FUNCTION FC 911 : VOID
TITLE =NEW FC911 (was FC1011) - Conveyors - Clearing Function
//New Order Sequence
//v0.1 2026-11-19: hold released at clearing start (FP M283.4); S3.2 lamp steady
//while held / blinking when ready; S3.2 held 3s releases the hold (T140).
//v0.2 2026-11-19: C10 empty proof added up over several runs (MD284), time from
//Surface_Length_10 (no more waiting for the bottomer). T137 no longer used.
//v0.3 2026-11-19: C10 empty proof by ENCODER TRAVEL (PIW 334 direct), not time:
//travel >= Surface_Length_10 + 20 % with exit clear, added up (MD284, MW288).
//v0.4 2026-11-19: encoder steps < 0 or > 300 pulses/scan ignored (Ch5 restarts
//from 0 when its gate reopens, every 500 mS while clearing) - no false proof.
NAME : CLEARING
VERSION : 0.4


VAR_TEMP
  EMPTY_11 : BOOL ;	//Empty Conveyor 11
  EMPTY_21 : BOOL ;	//Empty Conveyor 21
  EMPTY_12_22 : BOOL ;	//Empty Conveyor 12 & 22
  EMPTY_13_23 : BOOL ;	//Empty Conveyor 13 & 23
  C10_EMPTY_TEST : BOOL ;
  CLEARING_ABORT : BOOL ;
  PROOF_P : DINT ;	//C10 Empty Proof Travel [Pulses]
  D_ENC : DINT ;	//Encoder Pulses This Scan
  ENC_W : INT ;	//Encoder Word PIW 334
END_VAR
BEGIN
NETWORK
TITLE =HMI Clearing Call

      A     "M 140.3";
      A     "HMI_DB".CLEARING_SSW_MAIN;
      =     "M 5.2";
//;
      L     8;
      A     "M 10.0";
      =     "HMI_DB".CLEARING_SSW_STATUS;
      JC    CLEA;

      L     0;

CLEA: T     "HMI_DB".CLEARING_FUNCTION;

      A     "M 10.0";
      FN    "FN 155.7";
      R     "HMI_DB".CLEARING_SSW_MAIN;
      R     "M 54.2";
//;
      A     "M 5.2";
      FP    "FP 147.4";
      AN    "B 10.7"; // C11 - Empty
      AN    "B 11.0"; // C12 - Empty
      AN    "B 11.1"; // C13 - Empty
      AN    "B 11.2"; // C13 - Empty
      AN    "B 15.4"; // C21 - Empty
      AN    "B 15.5"; // C22 - Empty
      AN    "B 15.6"; // C23 - Empty
      AN    "B 15.7"; // C23 - Empty
      S     "M 54.2"; // Empty C11...C23
NETWORK
TITLE =New Order Seq - First New Order Packet to Pivot Conveyor 10
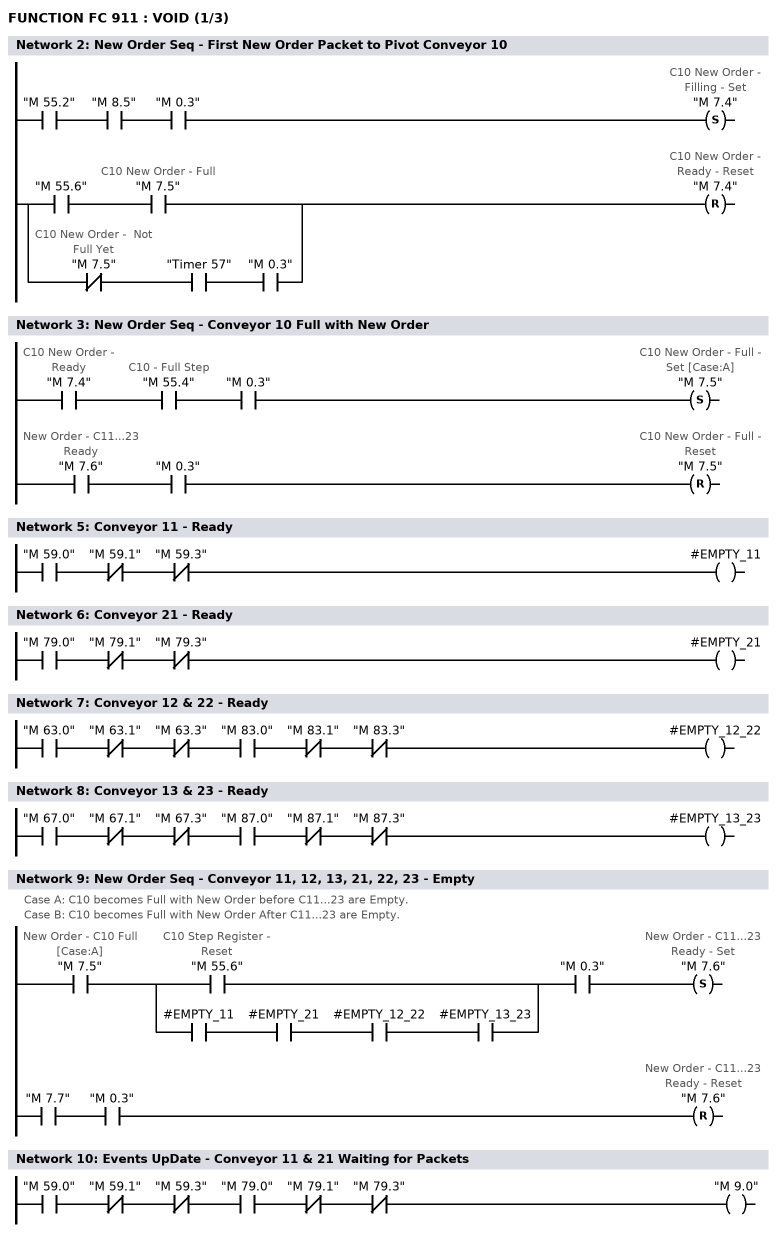

      A     "M 55.2";
      A     "M 8.5";
      A     "M 0.3";
      S     "M 7.4"; // C10 New Order - Filling - Set
//;
      A(    ;
      A     "M 55.6";
      A     "M 7.5"; // C10 New Order - Full
      O     ;
      AN    "M 7.5"; // C10 New Order -  Not Full Yet
      A     "Timer 57";
      A     "M 0.3";
      )     ;
      R     "M 7.4"; // C10 New Order - Ready - Reset
NETWORK
TITLE =New Order Seq - Conveyor 10 Full with New Order

      A     "M 7.4"; // C10 New Order - Ready
      A     "M 55.4"; // C10 - Full Step
      A     "M 0.3";
      S     "M 7.5"; // C10 New Order - Full - Set [Case:A]
//;
      A     "M 7.6"; // New Order - C11...23 Ready
      A     "M 0.3";
      R     "M 7.5"; // C10 New Order - Full - Reset
NETWORK
TITLE =New Order Seq
//New Order Seq - Waiting for the last Order Packets to Run out !


NETWORK
TITLE =Conveyor 11 - Ready

      A     "M 59.0";
      AN    "M 59.1";
      AN    "M 59.3";
      =     #EMPTY_11;
NETWORK
TITLE =Conveyor 21 - Ready

      A     "M 79.0";
      AN    "M 79.1";
      AN    "M 79.3";
      =     #EMPTY_21;
NETWORK
TITLE =Conveyor 12 & 22 - Ready

      A     "M 63.0";
      AN    "M 63.1";
      AN    "M 63.3";
      A     "M 83.0";
      AN    "M 83.1";
      AN    "M 83.3";
      =     #EMPTY_12_22;
NETWORK
TITLE =Conveyor 13 & 23 - Ready

      A     "M 67.0";
      AN    "M 67.1";
      AN    "M 67.3";
      A     "M 87.0";
      AN    "M 87.1";
      AN    "M 87.3";
      =     #EMPTY_13_23;
NETWORK
TITLE =New Order Seq - Conveyor 11, 12, 13, 21, 22, 23 - Empty
//Case A: C10 becomes Full with New Order before C11...23 are Empty.
//Case B: C10 becomes Full with New Order After C11...23 are Empty.
      A     "M 7.5"; // New Order - C10 Full [Case:A]
      A(    ;
      A     "M 55.6"; // C10 Step Register - Reset
      O     ;
      A     #EMPTY_11;
      A     #EMPTY_21;
      A     #EMPTY_12_22;
      A     #EMPTY_13_23;
      )     ;
      A     "M 0.3";
      S     "M 7.6"; // New Order - C11...23 Ready - Set
//;
      A     "M 7.7";
      A     "M 0.3";
      R     "M 7.6"; // New Order - C11...23 Ready - Reset
NETWORK
TITLE =Events UpDate - Conveyor 11 & 21 Waiting for Packets

      A     "M 59.0";
      AN    "M 59.1";
      AN    "M 59.3";
      A     "M 79.0";
      AN    "M 79.1";
      AN    "M 79.3";
      =     "M 9.0";
NETWORK
TITLE =New Order Seq - Conveyors 11, 21 - Empty
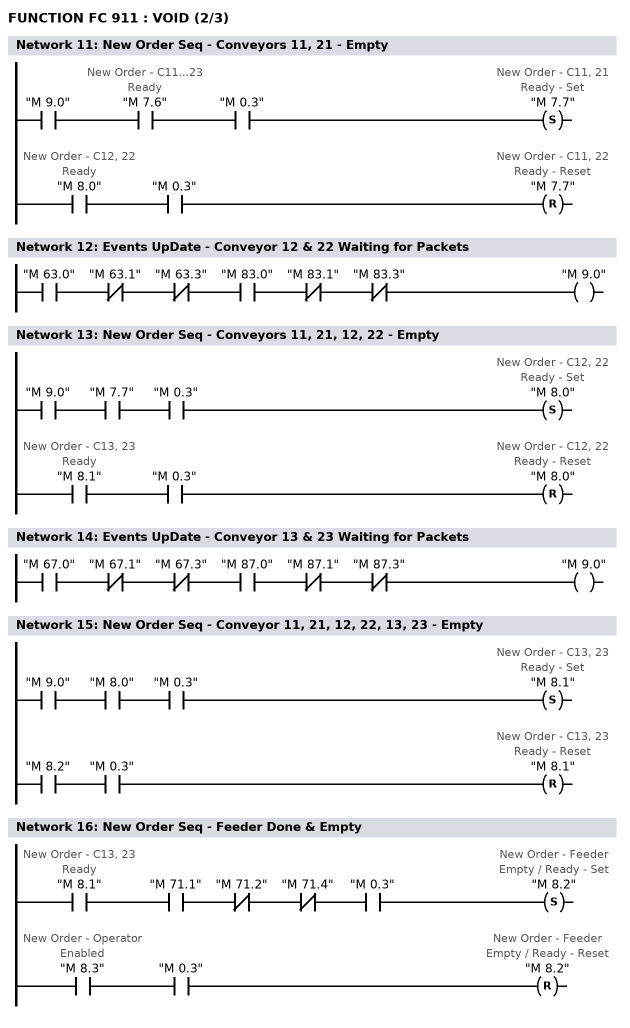

      A     "M 9.0";
      A     "M 7.6"; // New Order - C11...23 Ready
      A     "M 0.3";
      S     "M 7.7"; // New Order - C11, 21 Ready - Set
//;
      A     "M 8.0"; // New Order - C12, 22 Ready
      A     "M 0.3";
      R     "M 7.7"; // New Order - C11, 22 Ready - Reset
NETWORK
TITLE =Events UpDate - Conveyor 12 & 22 Waiting for Packets

      A     "M 63.0";
      AN    "M 63.1";
      AN    "M 63.3";
      A     "M 83.0";
      AN    "M 83.1";
      AN    "M 83.3";
      =     "M 9.0";
NETWORK
TITLE =New Order Seq - Conveyors 11, 21, 12, 22 - Empty

      A     "M 9.0";
      A     "M 7.7";
      A     "M 0.3";
      S     "M 8.0"; // New Order - C12, 22 Ready - Set
//;
      A     "M 8.1"; // New Order - C13, 23 Ready
      A     "M 0.3";
      R     "M 8.0"; // New Order - C12, 22 Ready - Reset
NETWORK
TITLE =Events UpDate - Conveyor 13 & 23 Waiting for Packets

      A     "M 67.0";
      AN    "M 67.1";
      AN    "M 67.3";
      A     "M 87.0";
      AN    "M 87.1";
      AN    "M 87.3";
      =     "M 9.0";
NETWORK
TITLE =New Order Seq - Conveyor 11, 21, 12, 22, 13, 23 - Empty

      A     "M 9.0";
      A     "M 8.0";
      A     "M 0.3";
      S     "M 8.1"; // New Order - C13, 23 Ready - Set
//;
      A     "M 8.2";
      A     "M 0.3";
      R     "M 8.1"; // New Order - C13, 23 Ready - Reset
NETWORK
TITLE =New Order Seq - Feeder Done & Empty

      A     "M 8.1"; // New Order - C13, 23 Ready
      A     "M 71.1";
      AN    "M 71.2";
      AN    "M 71.4";
      A     "M 0.3";
      S     "M 8.2"; // New Order - Feeder Empty / Ready - Set
//;
      A     "M 8.3"; // New Order - Operator Enabled
      A     "M 0.3";
      R     "M 8.2"; // New Order - Feeder Empty / Ready - Reset
NETWORK
TITLE =Conveyor 10 Clearing Enable after New Order
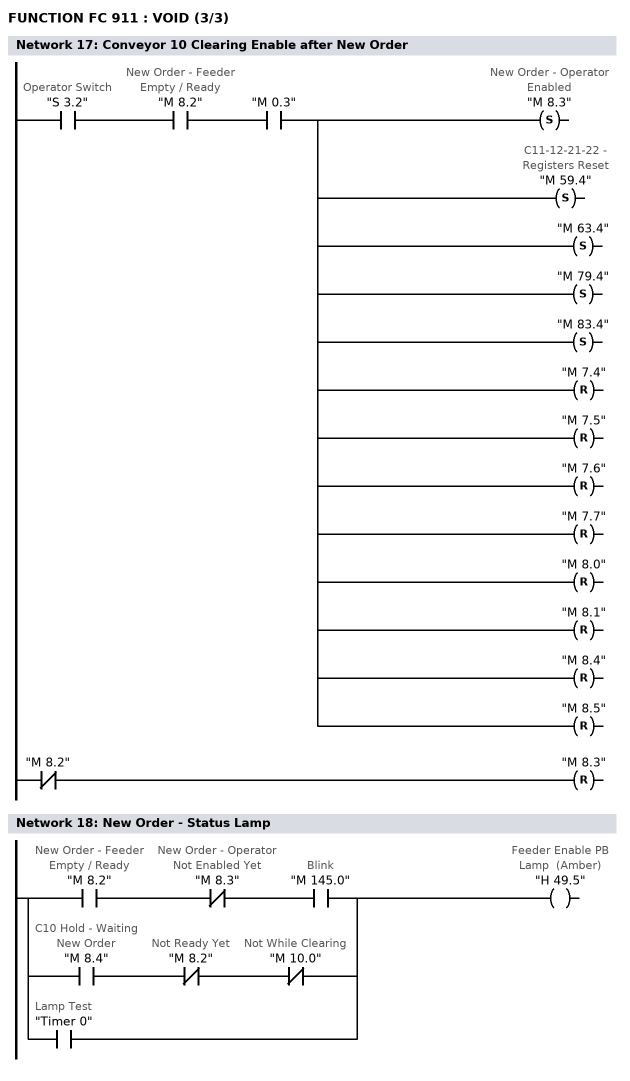

      A     "S 3.2"; // Operator Switch
      A     "M 8.2"; // New Order - Feeder Empty / Ready
      A     "M 0.3";
      S     "M 8.3"; // New Order - Operator Enabled
      S     "M 59.4"; // C11-12-21-22 - Registers Reset
      S     "M 63.4";
      S     "M 79.4";
      S     "M 83.4";
//;
      R     "M 7.4";
      R     "M 7.5";
      R     "M 7.6";
      R     "M 7.7";
      R     "M 8.0";
      R     "M 8.1";
      R     "M 8.4";
      R     "M 8.5";
//;
      ON    "M 8.2";
      R     "M 8.3";
NETWORK
TITLE =New Order - Status Lamp

//2026-11-19: BLINK = S3.2 can be pressed now (M8.2). STEADY = C10 held for the
//new order, not ready yet (M8.4 without M8.2) - before, the lamp stayed OFF.
      A(    ;
      A     "M 8.2"; // New Order - Feeder Empty / Ready
      AN    "M 8.3"; // New Order - Operator Not Enabled Yet
      A     "M 145.0"; // Blink
      )     ;
      O(    ;
      A     "M 8.4"; // C10 Hold - Waiting New Order
      AN    "M 8.2"; // Not Ready Yet
      AN    "M 10.0"; // Not While Clearing
      )     ;
      O     "Timer 0"; // Lamp Test
      =     "H 49.5"; // Feeder Enable PB Lamp  (Amber)
NETWORK
TITLE =S3.2 Held 3s - Release the Hold (Sequence Not Complete)
//2026-11-19: Before, S3.2 only worked with M8.2 (whole new-order chain done).
//If the chain got stuck, the TS waited with no way out but SIGNAL/F4.
//S3.2 held 3s releases the hold only (C11...C22 steps NOT reset: they may
//still carry the previous order).

      A     "S 3.2"; // Operator PB
      A     "M 8.4"; // C10 Hold Active
      AN    "M 10.0"; // Not While Clearing
      L     S5T#3S;
      SD    T    140; // Hold 3s (Free Timer)
//;
      A     T    140;
      A     "M 0.3";
      JCN   S321;

      R     "M 7.4";
      R     "M 7.5";
      R     "M 7.6";
      R     "M 7.7";
      R     "M 8.0";
      R     "M 8.1";
      R     "M 8.2";
      R     "M 8.3";
      R     "M 8.4"; // C10 Hold - Released
      R     "M 8.5"; // Clearing Done - Reset

S321: NOP   0;
NETWORK
TITLE =Conveyors Clearing Blink
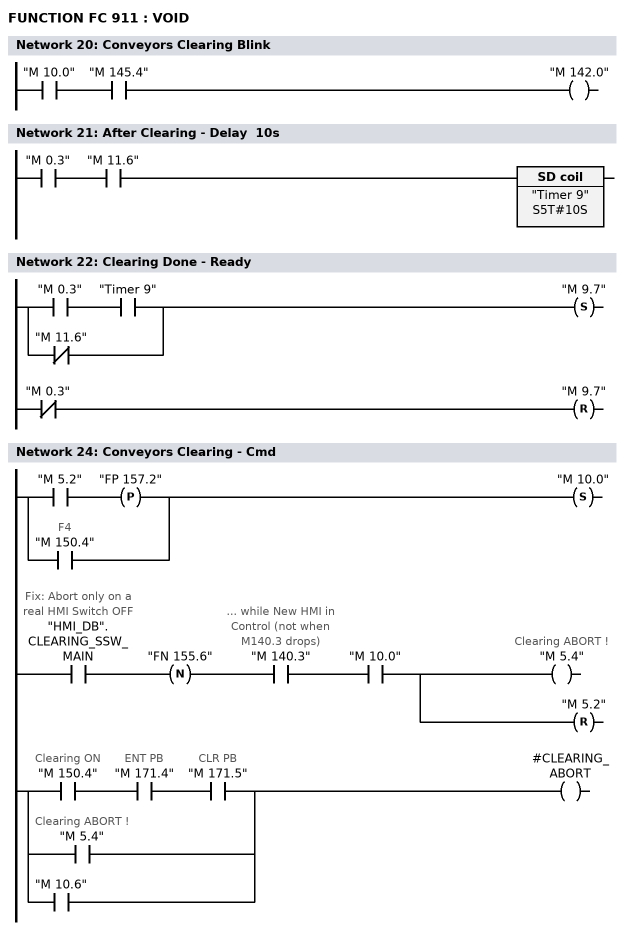

      A     "M 10.0";
      A     "M 145.4";
      =     "M 142.0";
NETWORK
TITLE =After Clearing - Delay  10s

      A     "M 0.3";
      A     "M 11.6";
      L     S5T#10S;
      SD    "Timer 9";
NETWORK
TITLE =Clearing Done - Ready

      A     "M 0.3";
      A     "Timer 9";
      ON    "M 11.6";
      S     "M 9.7";
//;
      ON    "M 0.3";
      R     "M 9.7";
NETWORK
TITLE =Clearing Command
//Clearing Command


NETWORK
TITLE =Conveyors Clearing - Cmd

      A(    ;
      A     "M 5.2";
      FP    "FP 157.2";
      O     ;
      A     "M 150.4"; // F4
      )     ;
      S     "M 10.0";
//;
      A     "HMI_DB".CLEARING_SSW_MAIN; // Fix: Abort only on a real HMI Switch OFF
      FN    "FN 155.6";
      A     "M 140.3"; // ... while New HMI in Control (not when M140.3 drops)
      A     "M 10.0";
      =     "M 5.4"; // Clearing ABORT !
      R     "M 5.2";
//;
      A(    ;
      A     "M 150.4"; // Clearing ON
      A     "M 171.4"; // ENT PB
      A     "M 171.5"; // CLR PB
      O     "M 5.4"; // Clearing ABORT !
      O     "M 10.6";
      )     ;
      =     #CLEARING_ABORT;
NETWORK
TITLE =Clearing Start - Release a Hold Left from the Previous Clearing
//Fix 2026-11-19: F4 pressed while C10 still held a new order (M8.4, S3.2 not
//pressed yet) -> C10 could not transfer, the clearing could never finish.
//F4 = clear everything: at every clearing start the hold and the new-order
//sequence are reset. They are set again when this clearing is done.

      A     "M 10.0"; // Clearing CMD
      FP    M    283.4; // Edge Memory (Free)
      JCN   CST1;

      R     "M 7.4";
      R     "M 7.5";
      R     "M 7.6";
      R     "M 7.7";
      R     "M 8.0";
      R     "M 8.1";
      R     "M 8.2";
      R     "M 8.3";
      R     "M 8.4"; // C10 Hold - Released
      R     "M 8.5"; // Clearing Done - Reset

CST1: NOP   0;
NETWORK
TITLE =Conveyors Clearing Conveyors 1,2,3,4 - TimeOut 30S
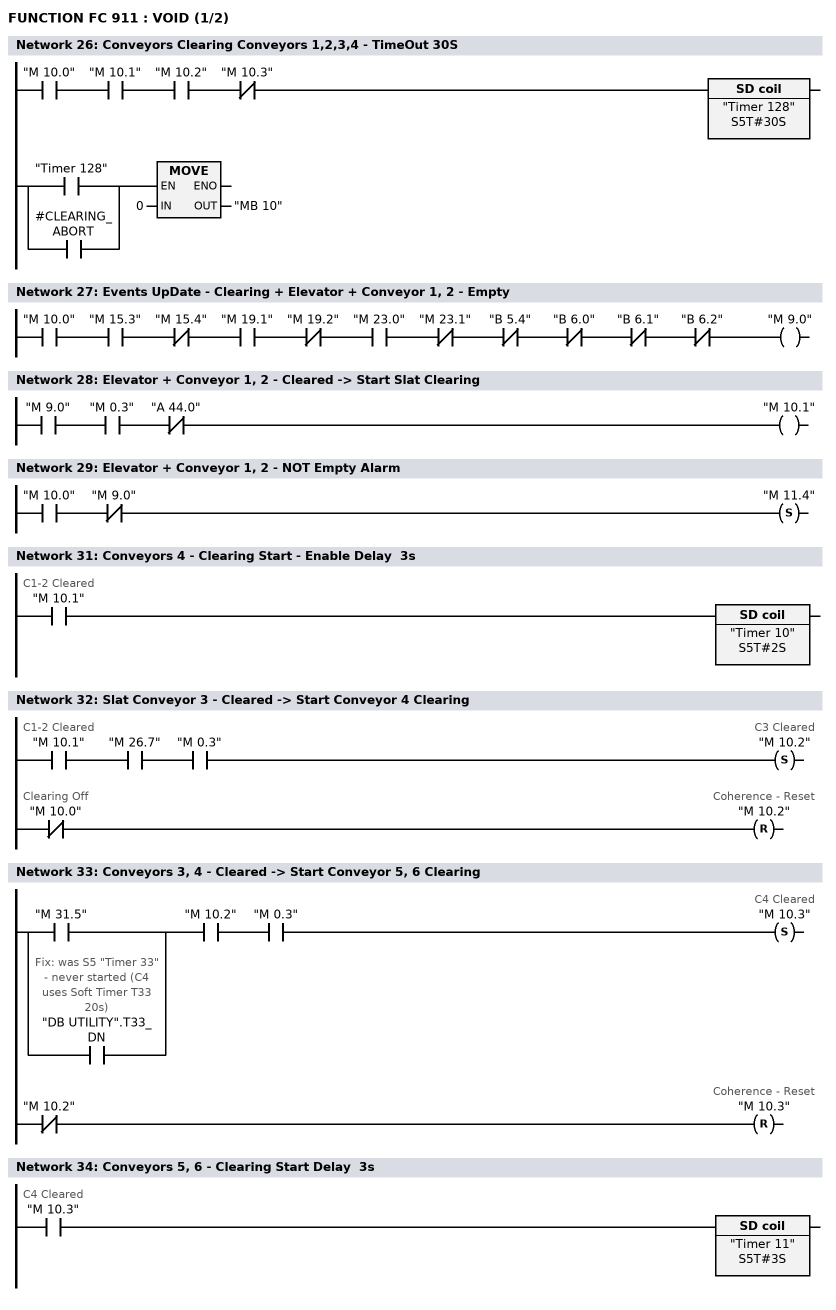

      A     "M 10.0";
      A     "M 10.1";
      A     "M 10.2";
      AN    "M 10.3";
      L     S5T#30S;
      SD    "Timer 128";
//;
      A     "Timer 128";
      O     #CLEARING_ABORT;
      JNB   NCLR;

      L     0;
      T     "MB 10"; // Clearing OFF

NCLR: NOP   0;
NETWORK
TITLE =Events UpDate - Clearing + Elevator + Conveyor 1, 2 - Empty

      A     "M 10.0";
      A     "M 15.3";
      AN    "M 15.4";
      A     "M 19.1";
      AN    "M 19.2";
      A     "M 23.0";
      AN    "M 23.1";
      AN    "B 5.4";
      AN    "B 6.0";
      AN    "B 6.1";
      AN    "B 6.2";
      =     "M 9.0";
NETWORK
TITLE =Elevator + Conveyor 1, 2 - Cleared -> Start Slat Clearing

      A     "M 9.0";
      A     "M 0.3";
      AN    "A 44.0";
      =     "M 10.1";
NETWORK
TITLE =Elevator + Conveyor 1, 2 - NOT Empty Alarm

      A     "M 10.0";
      AN    "M 9.0";
      S     "M 11.4";
NETWORK
TITLE =Clearing Sequence
//Clearing Sequence from Slat 3 to Pivot 10 Conveyors


NETWORK
TITLE =Conveyors 4 - Clearing Start - Enable Delay  3s

      A     "M 10.1"; // C1-2 Cleared
      L     S5T#2S;
      SD    "Timer 10";
NETWORK
TITLE =Slat Conveyor 3 - Cleared -> Start Conveyor 4 Clearing

      A     "M 10.1"; // C1-2 Cleared
      A     "M 26.7";
      A     "M 0.3";
      S     "M 10.2"; // C3 Cleared
//;
      AN    "M 10.0"; // Clearing Off
      R     "M 10.2"; // Coherence - Reset
NETWORK
TITLE =Conveyors 3, 4 - Cleared -> Start Conveyor 5, 6 Clearing

      A(    ;
      O     "M 31.5";
      O     "DB UTILITY".T33_DN; // Fix: was S5 "Timer 33" - never started (C4 uses Soft Timer T33 20s)
      )     ;
      A     "M 10.2";
      A     "M 0.3";
      S     "M 10.3"; // C4 Cleared
//;
      AN    "M 10.2";
      R     "M 10.3"; // Coherence - Reset
NETWORK
TITLE =Conveyors 5, 6 - Clearing Start Delay  3s

      A     "M 10.3"; // C4 Cleared
      L     S5T#3S;
      SD    "Timer 11"; // C4 Cleared Delayed
NETWORK
TITLE =Events UpDate - Conveyors 5, 6 - Clearing
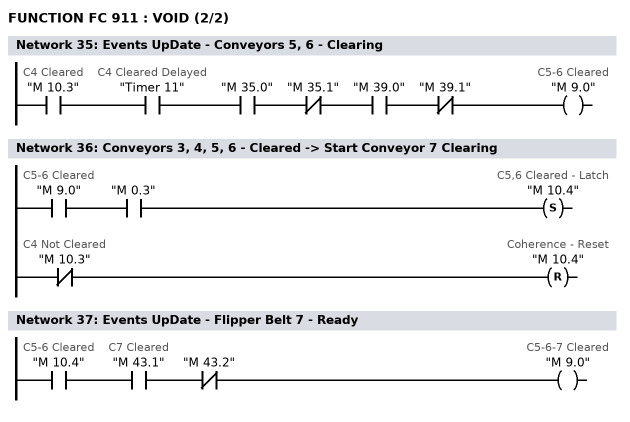

      A     "M 10.3"; // C4 Cleared
      A     "Timer 11"; // C4 Cleared Delayed
      A     "M 35.0";
      AN    "M 35.1";
      A     "M 39.0";
      AN    "M 39.1";
      =     "M 9.0"; // C5-6 Cleared
NETWORK
TITLE =Conveyors 3, 4, 5, 6 - Cleared -> Start Conveyor 7 Clearing

      A     "M 9.0"; // C5-6 Cleared
      A     "M 0.3";
      S     "M 10.4"; // C5,6 Cleared - Latch
//;
      AN    "M 10.3"; // C4 Not Cleared
      R     "M 10.4"; // Coherence - Reset
NETWORK
TITLE =Events UpDate - Flipper Belt 7 - Ready

      A     "M 10.4"; // C5-6 Cleared
      A     "M 43.1"; // C7 Cleared
      AN    "M 43.2";
      =     "M 9.0"; // C5-6-7 Cleared
NETWORK
TITLE =Conveyors 3, 4, 5, 6, 7, 8, 9 - Clearing - Cleared / Ready

      A     "M 9.0"; // C5-6-7 Cleared
      A     "M 47.2"; // C8 Cleared
      AN    "M 47.3";
      A     "M 51.1"; // C9 Cleared
      AN    "M 51.2";
      AN    "B 9.7"; // C9 - Pusher2 - Edge Cleared
      A     "M 0.3";
      L     S5T#3S;
      SD    "Timer 56"; // Delay 3s
//;
      A     "Timer 56";
      =     "M 10.5"; // C10 UpStream Cleared
      FP    "M 188.4";
      S     "M 58.2"; // C10 UpStream Cleared - Trigger Set
//;
      A     "M 10.5";
      L     S5T#1S;
      SE    "Timer 58"; // UpStream Cleared - Pulse 1s
NETWORK
TITLE =Clearing - C10 Proven Empty (Encoder Travel With Nothing Seen, Added Up)
//Fix: Clearing used to end with packets left on C10 (nothing checked C10 itself).
//v0.3 2026-11-19: proof by ENCODER TRAVEL, not time (C10 accelerates between
//B10.4 and B10.6). C10 encoder read directly every scan: PIW 334 = FM350-2 Ch5
//low word (HW Config 2026-11-19), wrap-safe difference per scan. Travel is
//ADDED UP over several runs (MD284) while the exit B10.6 is clear. Proven when
//travel >= C10 surface (Surface_Length_10, pulses) + 20 %. 0 -> 18000 p (5 m).
//Any packet seen on C10 (B10.3 / B10.4 / B10.5 / B10.6) or a Pusher 2 push
//restarts the proof (a pushed packet can sit at the infeed without C10 starting).

      L     "COLLATORS DB".Surface_Length_10; // C10 Surface [Pulses] (WORD)
      L     L#12;
      *D    ;
      L     L#10; // + 20 %
      /D    ;
      T     #PROOF_P;
//;
      L     #PROOF_P;
      L     L#1000;
      <D    ; // Surface Unknown (0) or Too Small
      JCN   P001;

      L     L#18000; // ~5 m @ 0.28 mm/pulse
      T     #PROOF_P;

P001: L     PIW  334; // C10 Encoder - Direct, Every Scan
      T     #ENC_W;
      A     "M 10.0"; // Clearing CMD
      JC    P002;

      L     #ENC_W; // No Clearing: Follow Encoder, Proof = 0
      T     MW   288;
      L     L#0;
      T     MD   284;
      JU    P004;

P002: L     #ENC_W; // Pulses Since Last Scan (INT Subtraction = Wrap-Safe)
      L     MW   288;
      -I    ;
      ITD   ;
      T     #D_ENC;
      L     #ENC_W;
      T     MW   288; // Last Encoder Word (Free)
      L     #D_ENC; // Counter Restart (Gate 5 Reopened, e.g. Every 500 mS in
      L     L#0; // Clearing) = Negative or Big Jump -> Not Travel: Ignore
      <D    ;
      JC    P006;

      L     #D_ENC;
      L     L#300; // Max Plausible Pulses per Scan
      >D    ;
      JCN   P003;

P006: L     L#0;
      T     #D_ENC;

P003: AN    "B 10.6"; // C10 Exit Sens Clear
      JCN   P004;

      L     MD   284; // Travel With Exit Clear, Added Up [Pulses] (Free)
      L     #D_ENC;
      +D    ;
      T     MD   284;

P004: A(    ;
      O     "B 10.3"; // Pusher Extended - Packet Sens (C10 Infeed)
      O     "M 51.7"; // Pusher 2 FWD - Packet Being Pushed
      O     "B 10.4"; // C10 InFeed Sens
      O     "B 10.5"; // C10 Full Sens
      O     "B 10.6"; // C10 Exit Sens
      )     ;
      JCN   P005;

      L     L#0; // Packet Seen - Proof Restarts
      T     MD   284;

P005: L     MD   284;
      L     #PROOF_P;
      >=D   ;
      A     "M 10.0";
      S     "M 10.7"; // C10 Proven Empty - Set
//;
      A(    ;
      O     "B 10.3";
      O     "M 51.7";
      O     "B 10.4";
      O     "B 10.5";
      O     "B 10.6";
      )     ;
      R     "M 10.7"; // Packet Seen - Not Empty
NETWORK
TITLE =Clearing - C10 Not Proven Empty -> Call C10 Transfer Again
//Fix: After a C10 transfer ends (C11/C21 full or 20s), packets could stay on C10
//and nothing called C10 again. While clearing and C10 is not proven empty,
//re-arm the C11/C21 call (M58.2) each time C10 is back to idle.
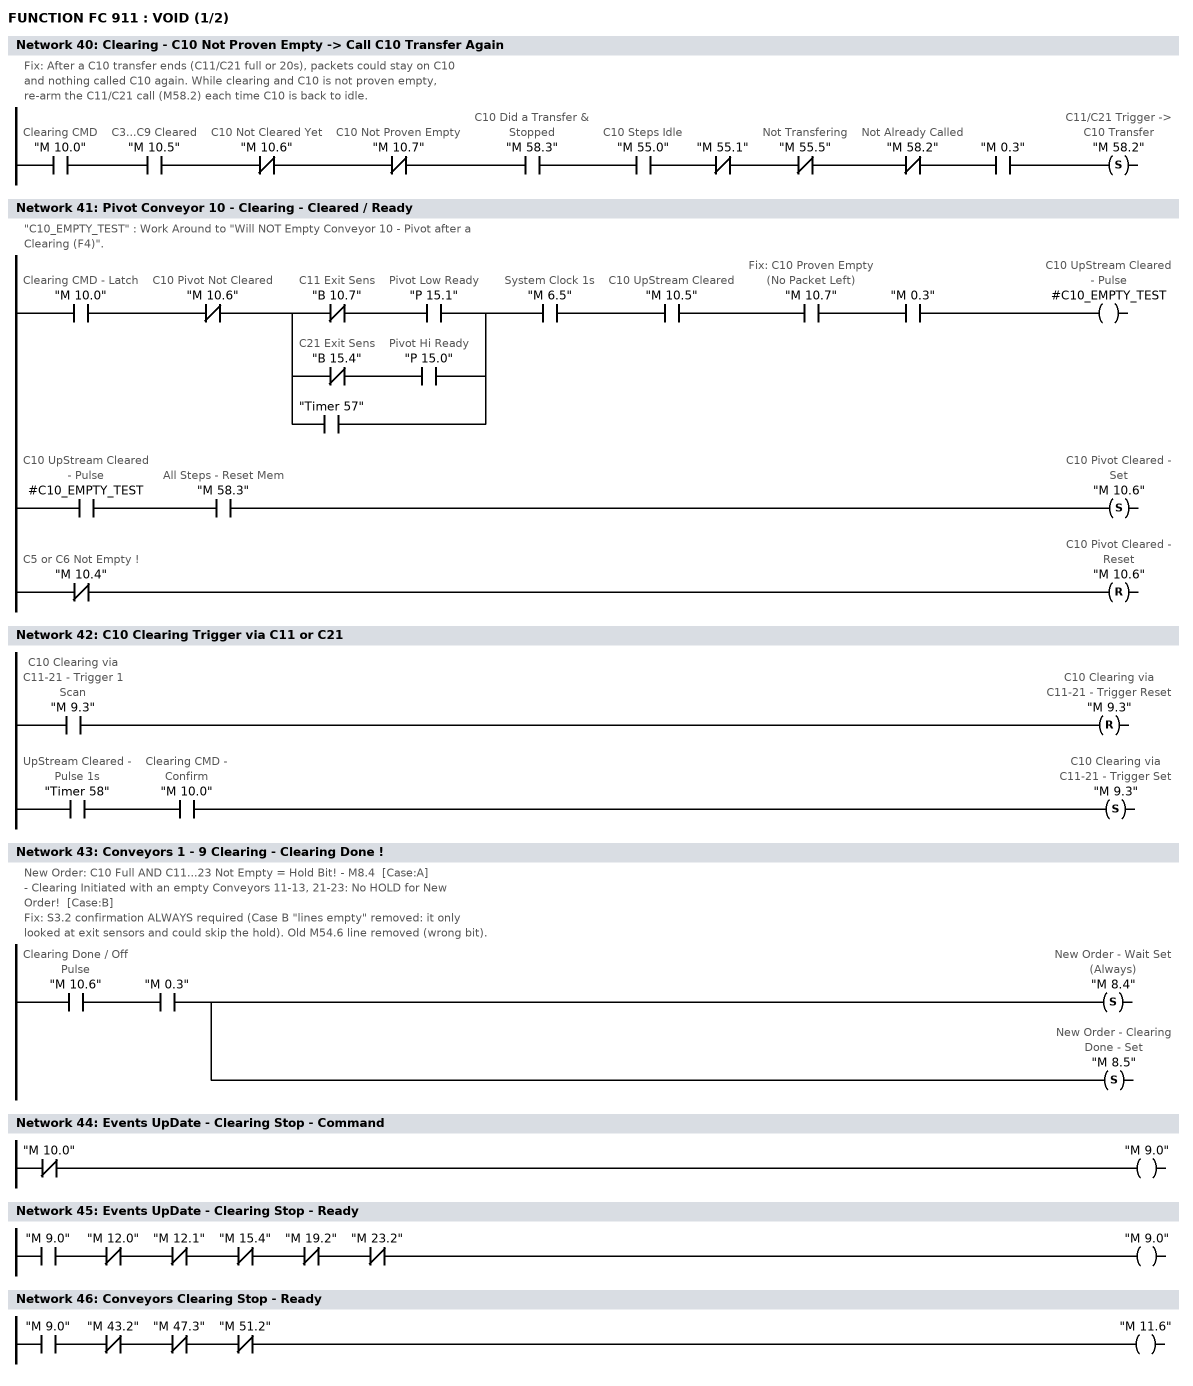
      A     "M 10.0"; // Clearing CMD
      A     "M 10.5"; // C3...C9 Cleared
      AN    "M 10.6"; // C10 Not Cleared Yet
      AN    "M 10.7"; // C10 Not Proven Empty
      A     "M 58.3"; // C10 Did a Transfer & Stopped
      A     "M 55.0"; // C10 Steps Idle
      AN    "M 55.1";
      AN    "M 55.5"; // Not Transfering
      AN    "M 58.2"; // Not Already Called
      A     "M 0.3";
      S     "M 58.2"; // C11/C21 Trigger -> C10 Transfer
NETWORK
TITLE =Pivot Conveyor 10 - Clearing - Cleared / Ready
//"C10_EMPTY_TEST" : Work Around to "Will NOT Empty Conveyor 10 - Pivot after a
//Clearing (F4)".
      A     "M 10.0"; // Clearing CMD - Latch
      AN    "M 10.6"; // C10 Pivot Not Cleared
      A(    ;
      AN    "B 10.7"; // C11 Exit Sens
      A     "P 15.1"; // Pivot Low Ready
      O     ;
      AN    "B 15.4"; // C21 Exit Sens
      A     "P 15.0"; // Pivot Hi Ready
      O     "Timer 57";
      )     ;
      A     "M 6.5"; // System Clock 1s
      A     "M 10.5"; // C10 UpStream Cleared
      A     "M 10.7"; // Fix: C10 Proven Empty (No Packet Left)
      A     "M 0.3";
      =     #C10_EMPTY_TEST; // C10 UpStream Cleared - Pulse
//;
      A     #C10_EMPTY_TEST; // C10 UpStream Cleared - Pulse
      A     "M 58.3"; // All Steps - Reset Mem
      S     "M 10.6"; // C10 Pivot Cleared - Set
//;
      AN    "M 10.4"; // C5 or C6 Not Empty !
      R     "M 10.6"; // C10 Pivot Cleared - Reset
NETWORK
TITLE =C10 Clearing Trigger via C11 or C21

      A     "M 9.3"; // C10 Clearing via C11-21 - Trigger 1 Scan
      R     "M 9.3"; // C10 Clearing via C11-21 - Trigger Reset
//;
      A     "Timer 58"; // UpStream Cleared - Pulse 1s
      A     "M 10.0"; // Clearing CMD - Confirm
      S     "M 9.3"; // C10 Clearing via C11-21 - Trigger Set
NETWORK
TITLE =Conveyors 1 - 9 Clearing - Clearing Done !
//New Order: C10 Full AND C11...23 Not Empty = Hold Bit! - M8.4  [Case:A]
//
//- Clearing Initiated with an empty Conveyors 11-13, 21-23: No HOLD for New
//Order!  [Case:B]
//
//Fix: S3.2 confirmation ALWAYS required (Case B "lines empty" removed: it only
//looked at exit sensors and could skip the hold). Old M54.6 line removed (wrong bit).
      A     "M 10.6"; // Clearing Done / Off Pulse
      A     "M 0.3";
      S     "M 8.4"; // New Order - Wait Set (Always)
      S     "M 8.5"; // New Order - Clearing Done - Set
NETWORK
TITLE =Events UpDate - Clearing Stop - Command

      AN    "M 10.0";
      =     "M 9.0";
NETWORK
TITLE =Events UpDate - Clearing Stop - Ready

      A     "M 9.0";
      AN    "M 12.0";
      AN    "M 12.1";
      AN    "M 15.4";
      AN    "M 19.2";
      AN    "M 23.2";
      =     "M 9.0";
NETWORK
TITLE =Conveyors Clearing Stop - Ready

      A     "M 9.0";
      AN    "M 43.2";
      AN    "M 47.3";
      AN    "M 51.2";
      =     "M 11.6";
NETWORK
TITLE =New Order
//New Order : Start Filling Conveyors


NETWORK
TITLE =Events UpDate - Elevator Packet IN
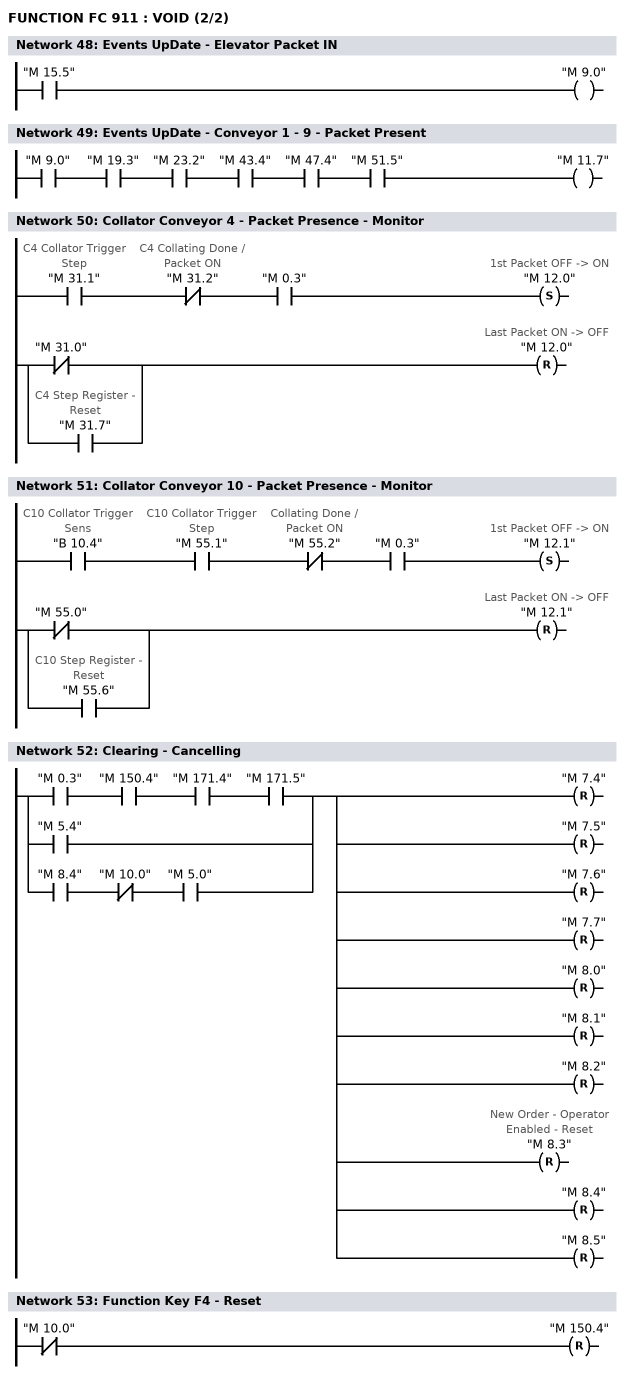

      A     "M 15.5";
      =     "M 9.0";
NETWORK
TITLE =Events UpDate - Conveyor 1 - 9 - Packet Present

      A     "M 9.0";
      A     "M 19.3";
      A     "M 23.2";
      A     "M 43.4";
      A     "M 47.4";
      A     "M 51.5";
      =     "M 11.7";
NETWORK
TITLE =Collator Conveyor 4 - Packet Presence - Monitor

      A     "M 31.1"; // C4 Collator Trigger Step
      AN    "M 31.2"; // C4 Collating Done / Packet ON
      A     "M 0.3";
      S     "M 12.0"; // 1st Packet OFF -> ON
//;
      A(    ;
      ON    "M 31.0";
      O     "M 31.7"; // C4 Step Register - Reset
      )     ;
      R     "M 12.0"; // Last Packet ON -> OFF
NETWORK
TITLE =Collator Conveyor 10 - Packet Presence - Monitor

      A     "B 10.4"; // C10 Collator Trigger Sens
      A     "M 55.1"; // C10 Collator Trigger Step
      AN    "M 55.2"; // Collating Done / Packet ON
      A     "M 0.3";
      S     "M 12.1"; // 1st Packet OFF -> ON
//;
      A(    ;
      ON    "M 55.0";
      O     "M 55.6"; // C10 Step Register - Reset
      )     ;
      R     "M 12.1"; // Last Packet ON -> OFF
NETWORK
TITLE =Clearing - Cancelling

      A     "M 0.3";
      A     "M 150.4";
      A     "M 171.4";
      A     "M 171.5";
      O     "M 5.4";
      O(    ;
      A     "M 8.4";
      AN    "M 10.0";
      A     "M 5.0";
      )     ;
      R     "M 7.4";
      R     "M 7.5";
      R     "M 7.6";
      R     "M 7.7";
      R     "M 8.0";
      R     "M 8.1";
      R     "M 8.2";
      R     "M 8.3"; // New Order - Operator Enabled - Reset
      R     "M 8.4";
      R     "M 8.5";
NETWORK
TITLE =Function Key F4 - Reset

      AN    "M 10.0";
      R     "M 150.4";
END_FUNCTION


FUNCTION FC 912 : VOID
TITLE =NEW FC912 (was FC1012) - Conveyor 0 & Pusher 0
NAME : 'Pos.1'
VERSION : 0.1


VAR_TEMP
  TIMER_RESET : BOOL ;
  MAIN_SERVICE_1_SW : BOOL ;
  CONV_0_SERVICE_FWD : BOOL ;
  CONV_0_SERVICE_REV : BOOL ;
  RESET_1 : BOOL ;
  RESET_2 : BOOL ;
  PUSHER_PUSH : BOOL ;
END_VAR
BEGIN
NETWORK
TITLE =Conveyor 0 - Service

      A     "HMI_DB".ALL_SERVICE_ENABLE_SW;
      A     "HMI_DB".CONVEYOR_0_SERVICE_SW;
      A     "HMI_DB".SERVICE_SW_1_STATUS;
      =     #MAIN_SERVICE_1_SW;
//;
      A     #MAIN_SERVICE_1_SW;
      O     "M 14.0";
      JNB   PUS0;
      A     "HMI_DB".HMI_ROLLER_TEST_FWD_SSW;
      FP    "FP 168.3";
      R     "HMI_DB".HMI_ROLLER_TEST_REV_SSW;
      =     #RESET_1;
//;
      A     "HMI_DB".HMI_ROLLER_TEST_REV_SSW;
      FP    "FP 168.4";
      R     "HMI_DB".HMI_ROLLER_TEST_FWD_SSW;
      =     #RESET_2;
//;
      A(    ;
      O     #RESET_1;
      O     #RESET_2;
      )     ;
      L     S5T#1S;
      SF    "Timer 110";
//;
      A     "HMI_DB".HMI_ROLLER_TEST_FWD_SSW;
      AN    "Timer 110";
      =     #CONV_0_SERVICE_FWD;
//;
      A     "HMI_DB".HMI_ROLLER_TEST_REV_SSW;
      AN    "Timer 110";
      =     #CONV_0_SERVICE_REV;
//;
      A     "HMI_DB".HMI_PUSHER_0_TEST_SSW;
      =     #PUSHER_PUSH;
//;
      AN    #MAIN_SERVICE_1_SW;
      R     "HMI_DB".HMI_ROLLER_TEST_FWD_SSW;
      R     "HMI_DB".HMI_ROLLER_TEST_REV_SSW;

PUS0: R     #CONV_0_SERVICE_FWD;
      R     #CONV_0_SERVICE_REV;
      R     #RESET_1;
      R     #RESET_2;
      R     #PUSHER_PUSH;
      FP    "FP 158.0";
      =     "M 14.0";
NETWORK
TITLE =Function Keys <F5 > on HMI - Reset
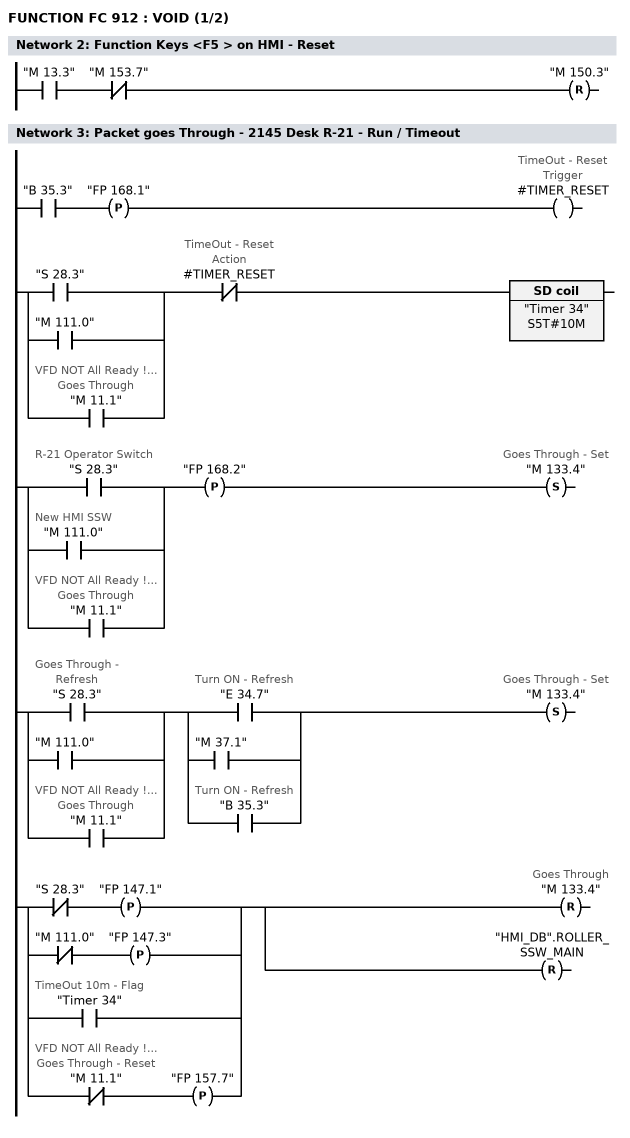

      A     "M 13.3";
      AN    "M 153.7";
      R     "M 150.3";
NETWORK
TITLE =Packet goes Through - 2145 Desk R-21 - Run / Timeout

      A     "B 35.3";
      FP    "FP 168.1";
      =     #TIMER_RESET; // TimeOut - Reset Trigger
//;
      A     "S 28.3";
      O     "M 111.0";
      O     "M 11.1"; // VFD NOT All Ready !... Goes Through
      AN    #TIMER_RESET; // TimeOut - Reset Action
      L     S5T#10M;
      SD    "Timer 34"; // TimeOut 10m
//;
      A     "S 28.3"; // R-21 Operator Switch
      O     "M 111.0"; // New HMI SSW
      O     "M 11.1"; // VFD NOT All Ready !... Goes Through
      FP    "FP 168.2"; // Turn ON - Pulse
      S     "M 133.4"; // Goes Through - Set
//;
      A     "S 28.3"; // Goes Through - Refresh
      O     "M 111.0";
      O     "M 11.1"; // VFD NOT All Ready !... Goes Through
      A(    ;
      O     "E 34.7"; // Turn ON - Refresh
      O     "M 37.1";
      O     "B 35.3"; // Turn ON - Refresh
      )     ;
      S     "M 133.4"; // Goes Through - Set
//;
      A(    ;
      O(    ;
      AN    "S 28.3";
      FP    "FP 147.1"; // Turn OFF - Pulse
      )     ;
      O(    ;
      AN    "M 111.0";
      FP    "FP 147.3"; // Turn OFF - Pulse
      O     "Timer 34"; // TimeOut 10m - Flag
      )     ;
      O(    ;
      AN    "M 11.1"; // VFD NOT All Ready !... Goes Through - Reset
      FP    "FP 157.7";
      )     ;
      )     ;
      R     "M 133.4"; // Goes Through
      R     "HMI_DB".ROLLER_SSW_MAIN;
NETWORK
TITLE =
//
//      A     "E 2.4"
//      S     "M 33.0"                    // Solid Detected ?
////;
//      A     "M 33.0"                    // Delay Timer - Start
//      L     S5T#300MS
//      SD    "Timer 26"                  // Debouncer 300mS
////;
//      A     "Timer 26"                  // Delayed Test Pulse
//      AN    "E 2.4"                     // Foul Detection
//      R     "M 33.0"                    // Not Detected !
////;
//      A     "Timer 26"                  // Delayed Test Pulse
//      A     "M 33.0"                    // Detection Comfirm !
//      =     "M 33.1"                    // Packet Height OK
//      R     "M 33.0"                    // Reset
//


NETWORK
TITLE =Packet Height - Sensing / Debouncing
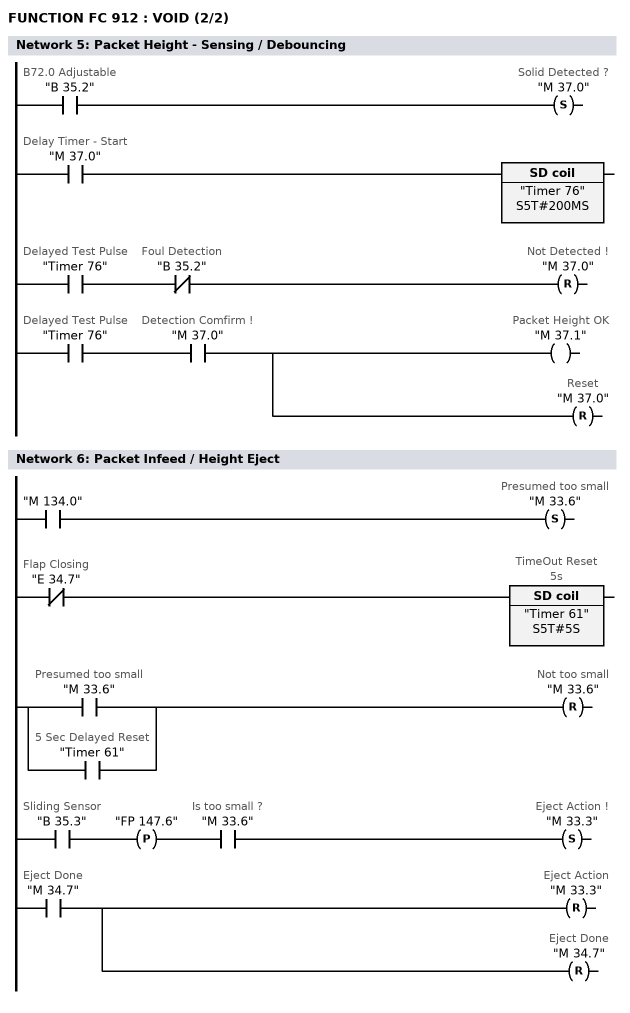

      A     "B 35.2"; // B72.0 Adjustable
      S     "M 37.0"; // Solid Detected ?
//;
      A     "M 37.0"; // Delay Timer - Start
      L     S5T#200MS;
      SD    "Timer 76"; // Debouncer 300mS
//;
      A     "Timer 76"; // Delayed Test Pulse
      AN    "B 35.2"; // Foul Detection
      R     "M 37.0"; // Not Detected !
//;
      A     "Timer 76"; // Delayed Test Pulse
      A     "M 37.0"; // Detection Comfirm !
      =     "M 37.1"; // Packet Height OK
      R     "M 37.0"; // Reset
NETWORK
TITLE =Packet Infeed / Height Eject

      A     "M 134.0";
      S     "M 33.6"; // Presumed too small
//;
      AN    "E 34.7"; // Flap Closing
      L     S5T#5S; // TimeOut Reset 5s
      SD    "Timer 61";
//;
      A     "M 33.6"; // Presumed too small
//    A     "M 33.1"                    // Packet Height OK ?
      O     "Timer 61"; // 5 Sec Delayed Reset
      R     "M 33.6"; // Not too small
//;
      A     "B 35.3"; // Sliding Sensor
      FP    "FP 147.6";
      A     "M 33.6"; // Is too small ?
      S     "M 33.3"; // Eject Action !
//;
      A     "M 34.7"; // Eject Done
      R     "M 33.3"; // Eject Action
      R     "M 34.7"; // Eject Done
NETWORK
TITLE =Eject Comfirmation

      A     "M 13.0";
      JNB   OUT1;

      A     "B 35.3";
      AN    "M 132.6"; // Not Triggered by Pusher
      S     "M 34.3"; // Eject Step 1
//;
      A     "B 35.4";
      AN    "M 132.6"; // Not Triggered by Pusher
      S     "M 34.4"; // Eject Step 2
//;
      A     "K 62.0"; // Conveyor 0 - Running
      A     "M 153.7";
      A     "M 34.3"; // Eject Step 1
      A     "M 34.4"; // Eject Step 2
      S     "M 34.5"; // Eject Step 3
//;
      A     "M 34.5"; // Eject Step 3
      AN    "B 35.4"; // Eject Step 4
      S     "M 34.7"; // Eject Done
      R     "M 34.3"; // Eject Step 1 - Reset
      R     "M 34.4"; // Eject Step 2 - Reset
      R     "M 34.5"; // Eject Step 3 - Reset
      R     "M 33.3"; // Eject Action - Reset
//;
      A     "M 132.5"; // Reset with Pusher Extend
      A     "B 35.4";
      R     "M 34.3"; // Eject Step 1 - Reset
      R     "M 34.4"; // Eject Step 2 - Reset
      R     "M 34.5"; // Eject Step 3 - Reset
      R     "M 33.3"; // Eject Action - Reset

OUT1: CLR   ;
NETWORK
TITLE =Packet goes Through - Conveyor 0 Man Run - LAUER F5
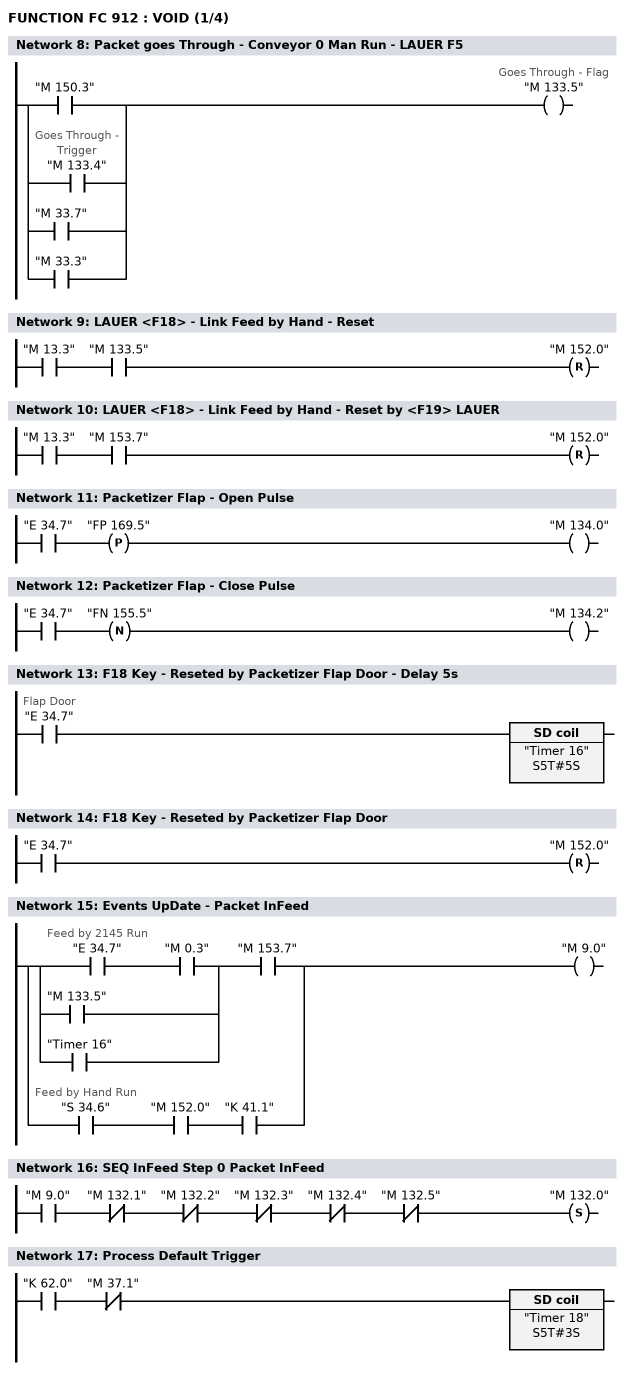

      O     "M 150.3";
      O     "M 133.4"; // Goes Through - Trigger
      O     "M 33.7";
      O     "M 33.3";
      =     "M 133.5"; // Goes Through - Flag
NETWORK
TITLE =LAUER <F18> - Link Feed by Hand - Reset

      A     "M 13.3";
      A     "M 133.5";
      R     "M 152.0";
NETWORK
TITLE =LAUER <F18> - Link Feed by Hand - Reset by <F19> LAUER

      A     "M 13.3";
      A     "M 153.7";
      R     "M 152.0";
NETWORK
TITLE =Packetizer Flap - Open Pulse

      A     "E 34.7";
      FP    "FP 169.5";
      =     "M 134.0";
NETWORK
TITLE =Packetizer Flap - Close Pulse

      A     "E 34.7";
      FN    "FN 155.5";
      =     "M 134.2";
NETWORK
TITLE =F18 Key - Reseted by Packetizer Flap Door - Delay 5s

      A     "E 34.7"; // Flap Door
      L     S5T#5S;
      SD    "Timer 16"; // Setup Mode Trigger
NETWORK
TITLE =F18 Key - Reseted by Packetizer Flap Door

      A     "E 34.7";
      R     "M 152.0";
NETWORK
TITLE =Events UpDate - Packet InFeed

      A(    ;
      A     "E 34.7"; // Feed by 2145 Run
      A     "M 0.3";
      O     "M 133.5";
      O     "Timer 16";
      A     "M 153.7";
      O     ;
      A     "S 34.6"; // Feed by Hand Run
      A     "M 152.0";
      A     "K 41.1";
      )     ;
      =     "M 9.0";
NETWORK
TITLE =SEQ InFeed Step 0 Packet InFeed

      A     "M 9.0";
      AN    "M 132.1";
      AN    "M 132.2";
      AN    "M 132.3";
      AN    "M 132.4";
      AN    "M 132.5";
      S     "M 132.0";
NETWORK
TITLE =Process Default Trigger

      A     "K 62.0";
      AN    "M 37.1";
      L     S5T#3S;
      SD    "Timer 18";
NETWORK
TITLE =Events UpDate
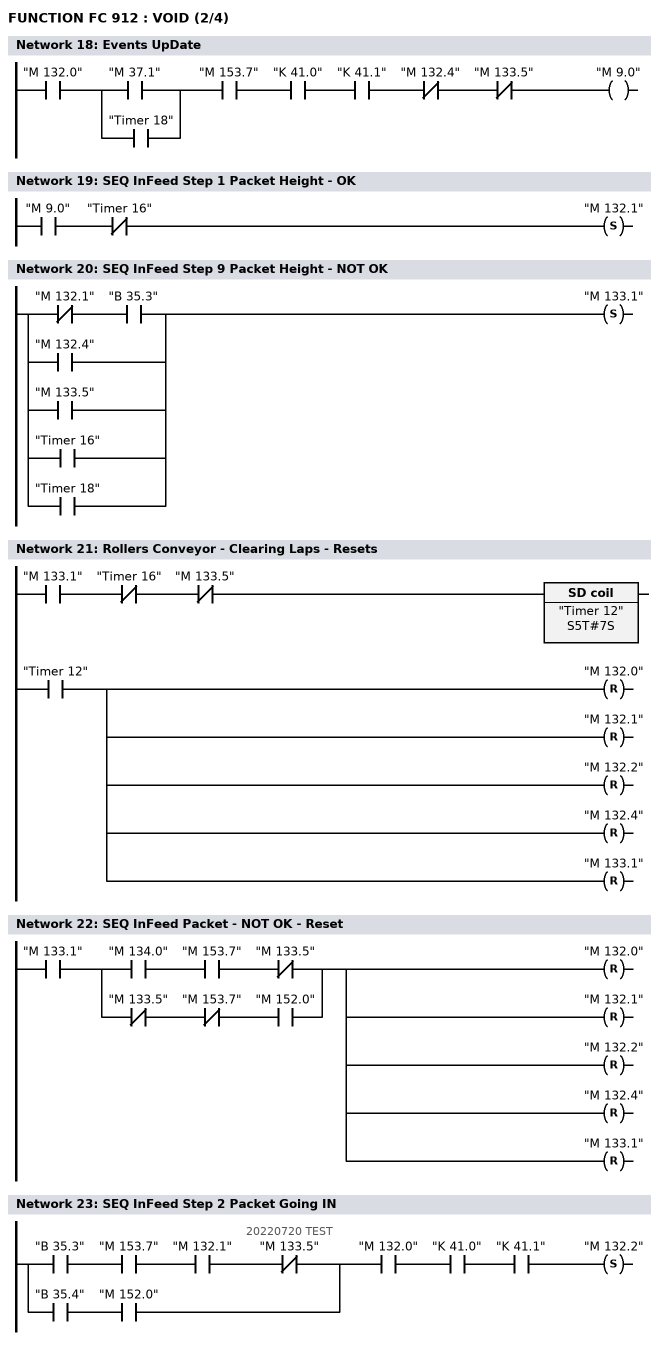

      A     "M 132.0";
      A(    ;
      O     "M 37.1";
      O     "Timer 18";
      )     ;
      A     "M 153.7";
      A     "K 41.0";
      A     "K 41.1";
      AN    "M 132.4";
      AN    "M 133.5";
      =     "M 9.0";
NETWORK
TITLE =SEQ InFeed Step 1 Packet Height - OK

      A     "M 9.0";
      AN    "Timer 16";
      S     "M 132.1";
NETWORK
TITLE =SEQ InFeed Step 9 Packet Height - NOT OK

      AN    "M 132.1";
      A     "B 35.3";
      O     "M 132.4";
      O     "M 133.5";
      O     "Timer 16";
      O     "Timer 18";
      S     "M 133.1";
NETWORK
TITLE =Rollers Conveyor - Clearing Laps - Resets

      A     "M 133.1";
      AN    "Timer 16";
      AN    "M 133.5";
      L     S5T#7S;
      SD    "Timer 12";
//;
      A     "Timer 12";
      R     "M 132.0";
      R     "M 132.1";
      R     "M 132.2";
      R     "M 132.4";
      R     "M 133.1";
NETWORK
TITLE =SEQ InFeed Packet - NOT OK - Reset

      A     "M 133.1";
      A(    ;
      A     "M 134.0";
      A     "M 153.7";
      AN    "M 133.5";
      O     ;
      AN    "M 133.5";
      AN    "M 153.7";
      A     "M 152.0";
      )     ;
      R     "M 132.0";
      R     "M 132.1";
      R     "M 132.2";
      R     "M 132.4";
      R     "M 133.1";
NETWORK
TITLE =SEQ InFeed Step 2 Packet Going IN

      A(    ;
      A     "B 35.3";
      A     "M 153.7";
      A     "M 132.1";
      AN    "M 133.5"; // 20220720 TEST
      O     ;
      A     "B 35.4";
      A     "M 152.0";
      )     ;
      A     "M 132.0";
      A     "K 41.0";
      A     "K 41.1";
      S     "M 132.2";
NETWORK
TITLE =SEQ InFeed Step 3 Conveyor Stop
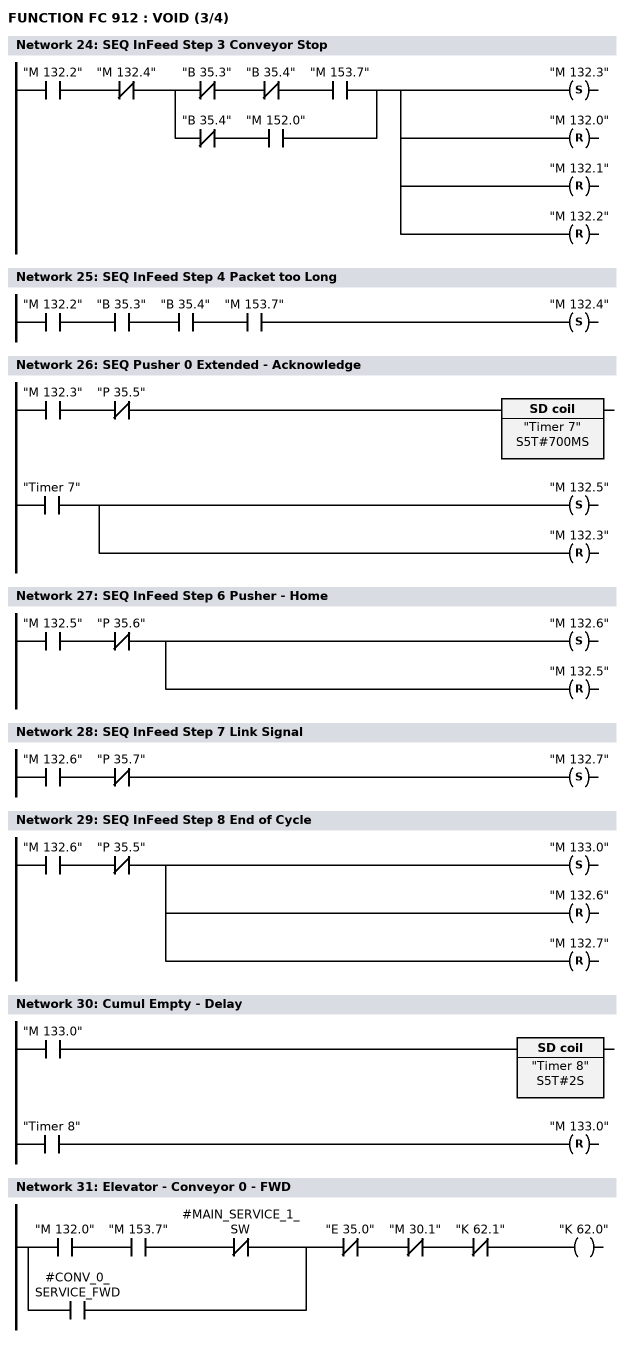

      A     "M 132.2";
      AN    "M 132.4";
      A(    ;
      AN    "B 35.3";
      AN    "B 35.4";
      A     "M 153.7";
      O     ;
      AN    "B 35.4";
      A     "M 152.0";
      )     ;
      S     "M 132.3";
      R     "M 132.0";
      R     "M 132.1";
      R     "M 132.2";
NETWORK
TITLE =SEQ InFeed Step 4 Packet too Long

      A     "M 132.2";
      A     "B 35.3";
      A     "B 35.4";
      A     "M 153.7";
      S     "M 132.4";
NETWORK
TITLE =SEQ Pusher 0 Extended - Acknowledge

      A     "M 132.3";
      AN    "P 35.5";
      L     S5T#700MS;
      SD    "Timer 7";
//;
      A     "Timer 7";
      S     "M 132.5";
      R     "M 132.3";
NETWORK
TITLE =SEQ InFeed Step 6 Pusher - Home

      A     "M 132.5";
      AN    "P 35.6";
      S     "M 132.6";
      R     "M 132.5";
NETWORK
TITLE =SEQ InFeed Step 7 Link Signal

      A     "M 132.6";
      AN    "P 35.7";
      S     "M 132.7";
NETWORK
TITLE =SEQ InFeed Step 8 End of Cycle

      A     "M 132.6";
      AN    "P 35.5";
      S     "M 133.0";
      R     "M 132.6";
      R     "M 132.7";
NETWORK
TITLE =Cumul Empty - Delay

      A     "M 133.0";
      L     S5T#2S;
      SD    "Timer 8";
//;
      A     "Timer 8";
      R     "M 133.0";
NETWORK
TITLE =Elevator - Conveyor 0 - FWD

      A(    ;
      A     "M 132.0";
      A     "M 153.7";
      AN    #MAIN_SERVICE_1_SW;
      O     #CONV_0_SERVICE_FWD;
      )     ;
      AN    "E 35.0";
      AN    "M 30.1";
      AN    "K 62.1";
      =     "K 62.0";
NETWORK
TITLE =Elevator - Conveyor 0 - REV
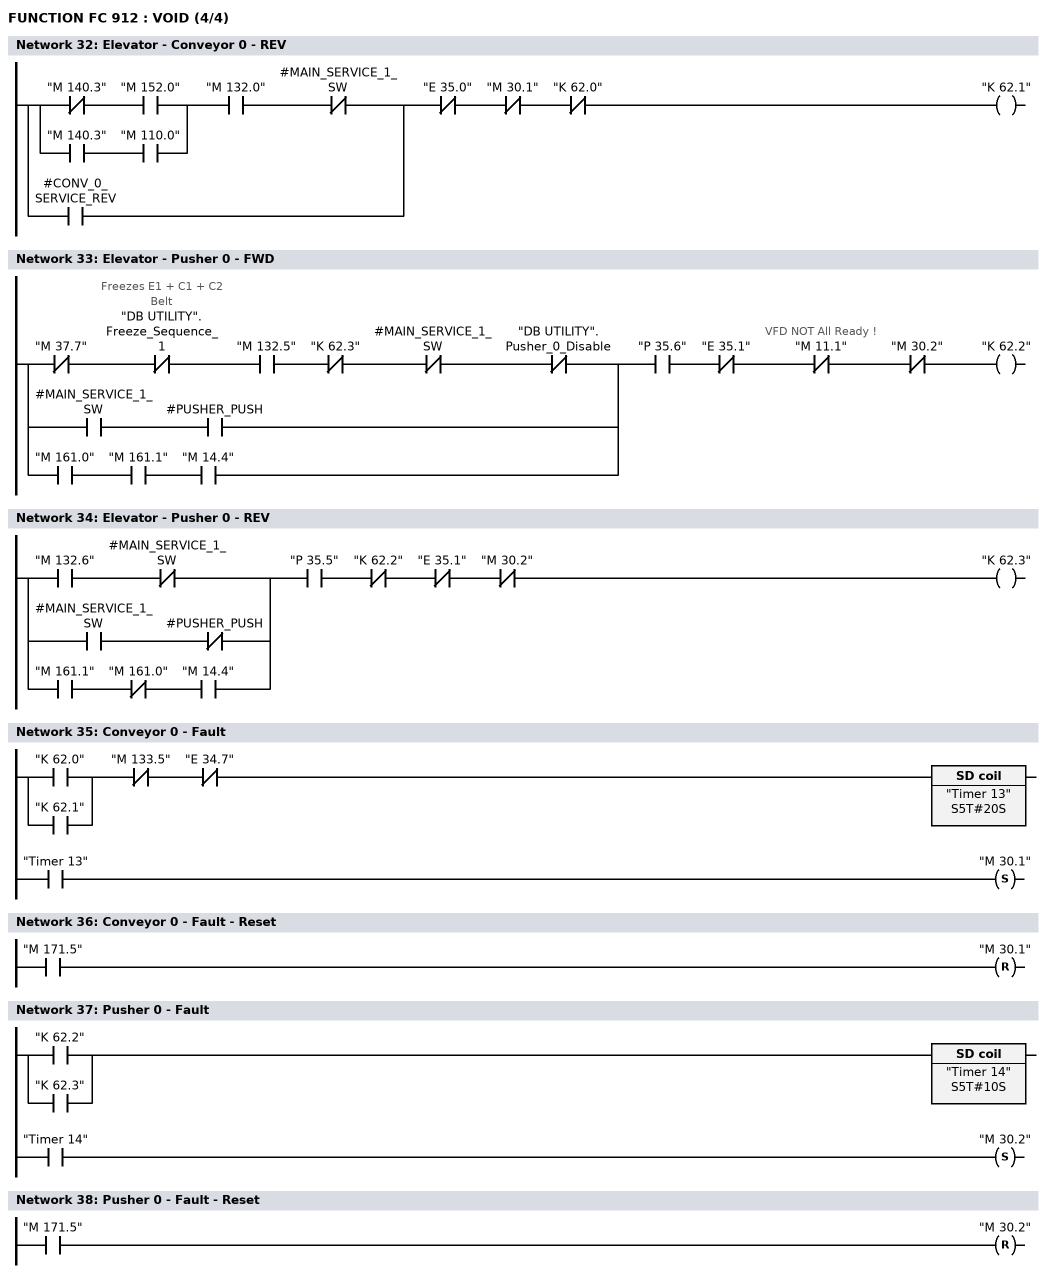

      A(    ;
      A(    ;
      AN    "M 140.3";
      A     "M 152.0";
      O     ;
      A     "M 140.3";
      A     "M 110.0";
      )     ;
      A     "M 132.0";
//     A     "M 152.0"
      AN    #MAIN_SERVICE_1_SW;
      O     #CONV_0_SERVICE_REV;
      )     ;
      AN    "E 35.0";
      AN    "M 30.1";
      AN    "K 62.0";
      =     "K 62.1";
NETWORK
TITLE =Elevator - Pusher 0 - FWD

      A(    ;
      AN    "M 37.7";
      AN    "DB UTILITY".Freeze_Sequence_1; //  Freezes E1 + C1 + C2 Belt
      A     "M 132.5";
      AN    "K 62.3";
      AN    #MAIN_SERVICE_1_SW;
      AN    "DB UTILITY".Pusher_0_Disable;
      O(    ;
      A     #MAIN_SERVICE_1_SW;
      A     #PUSHER_PUSH;
      )     ;
      O     ;
      A     "M 161.0";
      A     "M 161.1";
      A     "M 14.4";
      )     ;
      A     "P 35.6";
      AN    "E 35.1";
      AN    "M 11.1"; // VFD NOT All Ready !
      AN    "M 30.2";
      =     "K 62.2";
NETWORK
TITLE =Elevator - Pusher 0 - REV

      A(    ;
      A     "M 132.6";
      AN    #MAIN_SERVICE_1_SW;
      O(    ;
      A     #MAIN_SERVICE_1_SW;
      AN    #PUSHER_PUSH;
      )     ;
      O     ;
      A     "M 161.1";
      AN    "M 161.0";
      A     "M 14.4";
      )     ;
      A     "P 35.5";
      AN    "K 62.2";
      AN    "E 35.1";
      AN    "M 30.2";
      =     "K 62.3";
NETWORK
TITLE =Conveyor 0 - Fault

      A(    ;
      O     "K 62.0";
      O     "K 62.1";
      )     ;
      AN    "M 133.5";
      AN    "E 34.7";
      L     S5T#20S;
      SD    "Timer 13";
//;
      A     "Timer 13";
      S     "M 30.1";
NETWORK
TITLE =Conveyor 0 - Fault - Reset

      A     "M 171.5";
      R     "M 30.1";
NETWORK
TITLE =Pusher 0 - Fault

      A(    ;
      O     "K 62.2";
      O     "K 62.3";
      )     ;
      L     S5T#10S;
      SD    "Timer 14";
//;
      A     "Timer 14";
      S     "M 30.2";
NETWORK
TITLE =Pusher 0 - Fault - Reset

      A     "M 171.5";
      R     "M 30.2";
END_FUNCTION


FUNCTION FC 916 : VOID
TITLE =NEW FC916 (was FC1016) - Elevator + Pusher 1 Pos.2
//
NAME : POS_2
VERSION : 0.0


VAR_TEMP
  ELEVATOR_UP_OUT : BOOL ;
  ELEVATOR_DN_OUT : BOOL ;
  MAIN_SERVICE_1_SW : BOOL ;
  ELEVATOR_SERVICE_SW : BOOL ;
  ELEVATOR_DN_PB : BOOL ;
  ELEVATOR_UP_PB : BOOL ;
  ELEVATOR_ROUNDTRIP : BOOL ;
  PUSHER_PUSH : BOOL ;
  INITIALISATION : BOOL ;
  BRAKE_RELEASE_OK : BOOL ;
  BRAKE_CONTACTOR_KO : BOOL ;
END_VAR
BEGIN
NETWORK
TITLE =Elevator - Health OK
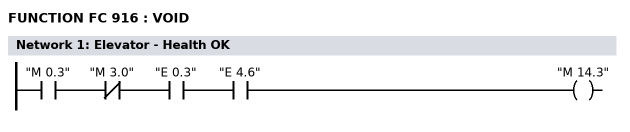

      A     "M 0.3";
      AN    "M 3.0";
      A     "E 0.3";
      A     "E 4.6";
      =     "M 14.3";
NETWORK
TITLE =Elevator - Service

      A     "HMI_DB".ALL_SERVICE_ENABLE_SW;
      A     "HMI_DB".ELEVATOR_SERVICE_SW;
      A     "HMI_DB".SERVICE_SW_1_STATUS;
      =     #MAIN_SERVICE_1_SW;
//;
      A     #MAIN_SERVICE_1_SW;
      O     "M 14.1";
      JNB   PUS1;
      A     "HMI_DB".HMI_ELEVATOR_SERVICE_SSW;
      =     #ELEVATOR_SERVICE_SW;
      S     "DB UTILITY".Pusher_0_Disable;
//;
      A     #ELEVATOR_SERVICE_SW;
      A(    ;
      A     "HMI_DB".HMI_ELEVATOR_TEST_DN_SSW;
      )     ;
      =     #ELEVATOR_DN_PB;
//;
      A     #ELEVATOR_SERVICE_SW;
      A(    ;
      A     "HMI_DB".HMI_ELEVATOR_TEST_UP_SSW;
      )     ;
      =     #ELEVATOR_UP_PB;
//;
      A     #MAIN_SERVICE_1_SW;
      AN    #ELEVATOR_SERVICE_SW;
      A     "HMI_DB".ELEVATOR_ROUND_TRIP_SSW;
      =     #ELEVATOR_ROUNDTRIP;
//;
      A     "HMI_DB".HMI_PUSHER_1_TEST_SSW;
      =     #PUSHER_PUSH;
//;
      AN    #MAIN_SERVICE_1_SW;
      R     "HMI_DB".HMI_ELEVATOR_SERVICE_SSW;
      R     "HMI_DB".HMI_ELEVATOR_TEST_DN_SSW;
      R     "HMI_DB".HMI_ELEVATOR_TEST_UP_SSW;
      R     "DB UTILITY".Pusher_0_Disable;

PUS1: R     #ELEVATOR_SERVICE_SW;
      R     #ELEVATOR_DN_PB;
      R     #ELEVATOR_UP_PB;
      R     #ELEVATOR_ROUNDTRIP;
      R     #PUSHER_PUSH;
      FP    "FP 158.1";
      =     "M 14.1";
//;
      A     "HMI_DB".SERVICE_INIT_PB;
      A     #ELEVATOR_SERVICE_SW;
      A     #MAIN_SERVICE_1_SW;
      =     #INITIALISATION;
NETWORK
TITLE =Elevator - Manual Run - Conditions
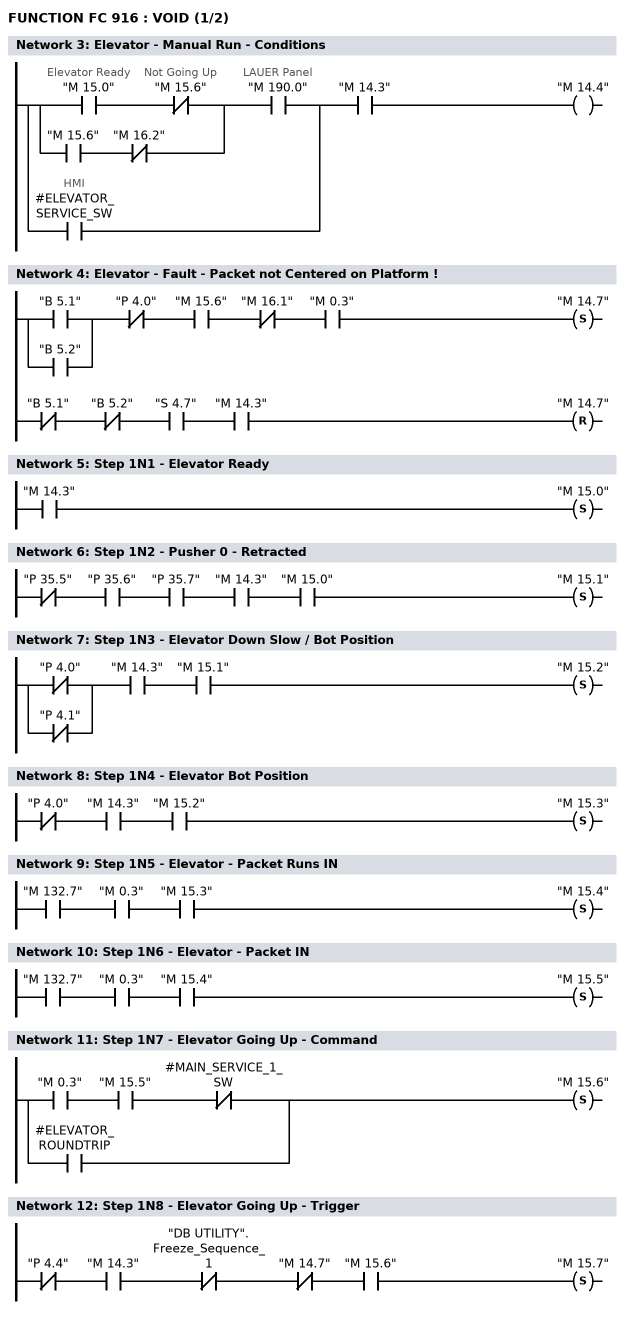

      A(    ;
      A     "M 15.0"; // Elevator Ready
      AN    "M 15.6"; // Not Going Up
      O     ; // or
      A     "M 15.6";
      AN    "M 16.2";
      )     ;
      A     "M 190.0"; // LAUER Panel
      O     #ELEVATOR_SERVICE_SW; // HMI
      A     "M 14.3";
      =     "M 14.4";
NETWORK
TITLE =Elevator - Fault - Packet not Centered on Platform !

      A(    ;
      O     "B 5.1";
      O     "B 5.2";
      )     ;
      AN    "P 4.0";
      A     "M 15.6";
      AN    "M 16.1";
      A     "M 0.3";
      S     "M 14.7";
//;
      AN    "B 5.1";
      AN    "B 5.2";
      A     "S 4.7";
      A     "M 14.3";
      R     "M 14.7";
NETWORK
TITLE =Step 1N1 - Elevator Ready

      A     "M 14.3";
      S     "M 15.0";
NETWORK
TITLE =Step 1N2 - Pusher 0 - Retracted

      AN    "P 35.5";
      A     "P 35.6";
      A     "P 35.7";
      A     "M 14.3";
      A     "M 15.0";
      S     "M 15.1";
NETWORK
TITLE =Step 1N3 - Elevator Down Slow / Bot Position

      A(    ;
      ON    "P 4.0";
      ON    "P 4.1";
      )     ;
      A     "M 14.3";
      A     "M 15.1";
      S     "M 15.2";
NETWORK
TITLE =Step 1N4 - Elevator Bot Position

      AN    "P 4.0";
      A     "M 14.3";
      A     "M 15.2";
      S     "M 15.3";
NETWORK
TITLE =Step 1N5 - Elevator - Packet Runs IN

      A     "M 132.7";
      A     "M 0.3";
      A     "M 15.3";
      S     "M 15.4";
NETWORK
TITLE =Step 1N6 - Elevator - Packet IN

      A     "M 132.7";
      A     "M 0.3";
      A     "M 15.4";
      S     "M 15.5";
NETWORK
TITLE =Step 1N7 - Elevator Going Up - Command

      A     "M 0.3";
      A     "M 15.5";
      AN    #MAIN_SERVICE_1_SW;
      O     #ELEVATOR_ROUNDTRIP;
      S     "M 15.6";
NETWORK
TITLE =Step 1N8 - Elevator Going Up - Trigger

      AN    "P 4.4";
      A     "M 14.3";
      AN    "DB UTILITY".Freeze_Sequence_1;
      AN    "M 14.7";
      A     "M 15.6";
      S     "M 15.7";
NETWORK
TITLE =Step 1N9 - Elevator Going Up - Slow
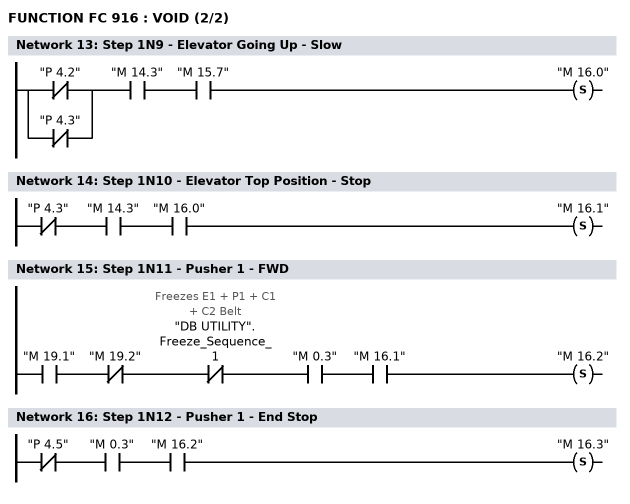

      A(    ;
      ON    "P 4.2";
      ON    "P 4.3";
      )     ;
      A     "M 14.3";
      A     "M 15.7";
      S     "M 16.0";
NETWORK
TITLE =Step 1N10 - Elevator Top Position - Stop

      AN    "P 4.3";
      A     "M 14.3";
      A     "M 16.0";
      S     "M 16.1";
NETWORK
TITLE =Step 1N11 - Pusher 1 - FWD

      A     "M 19.1";
      AN    "M 19.2";
      AN    "DB UTILITY".Freeze_Sequence_1; //  Freezes E1 + P1 + C1 + C2 Belt
      A     "M 0.3";
      A     "M 16.1";
      S     "M 16.2";
NETWORK
TITLE =Step 1N12 - Pusher 1 - End Stop

      AN    "P 4.5";
      A     "M 0.3";
      A     "M 16.2";
      S     "M 16.3";
NETWORK
TITLE =Soft Timer 15 Reset

      A     "M 16.3";
      AN    "M 16.4";
      A     "M 14.3";
      A     "M 0.3";
      JCN   R151;
      JU    E151;

R151: L     L#0;
      T     "DB UTILITY".T15_ET;
      R     "DB UTILITY".T15_DN;

E151: NOP   0;

NETWORK
TITLE =Soft Timer 15 Add

      A     "M 16.3";
      AN    "M 16.4";
      A     "M 14.3";
      A     "M 0.3";
      AN    "DB UTILITY".Freeze_Sequence_1;
      AN    "DB UTILITY".T15_DN;
      JCN   E152;

      L     "DB UTILITY".T15_ET;
      L     "DB UTILITY".Scan_Cycle_Previous;
      ITD   ;
      +D    ;
      T     "DB UTILITY".T15_ET;

E152: NOP   0;

NETWORK
TITLE =Soft Timer 15 Done 100mS
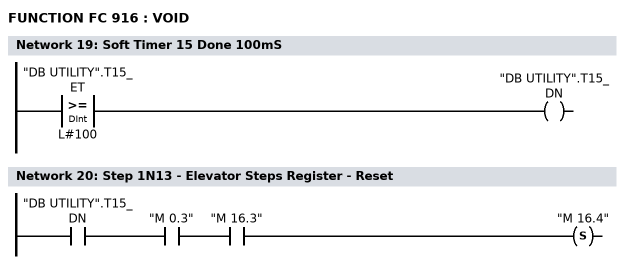

      L     "DB UTILITY".T15_ET;
      L     L#100;
      >=D   ;
      =     "DB UTILITY".T15_DN;

NETWORK
TITLE =Step 1N13 - Elevator Steps Register - Reset

      A     "DB UTILITY".T15_DN;
      A     "M 0.3";
      A     "M 16.3";
      S     "M 16.4";
NETWORK
TITLE =Elevator Steps Register - Reset

      A(    ;
      A     "M 190.0";
      A     "M 171.4";
      A     "M 171.5";
      O     "M 16.4";
      O     #INITIALISATION;
      O     "DB UTILITY".Elevator_Disable;
      )     ;
      A     "M 0.3";
      JC    M001;
      JU    M002;

M001: L     W#16#0;
      T     "MW 15";

M002: CLR   ;
NETWORK
TITLE =Trans System - Ready -> Tuber 2145
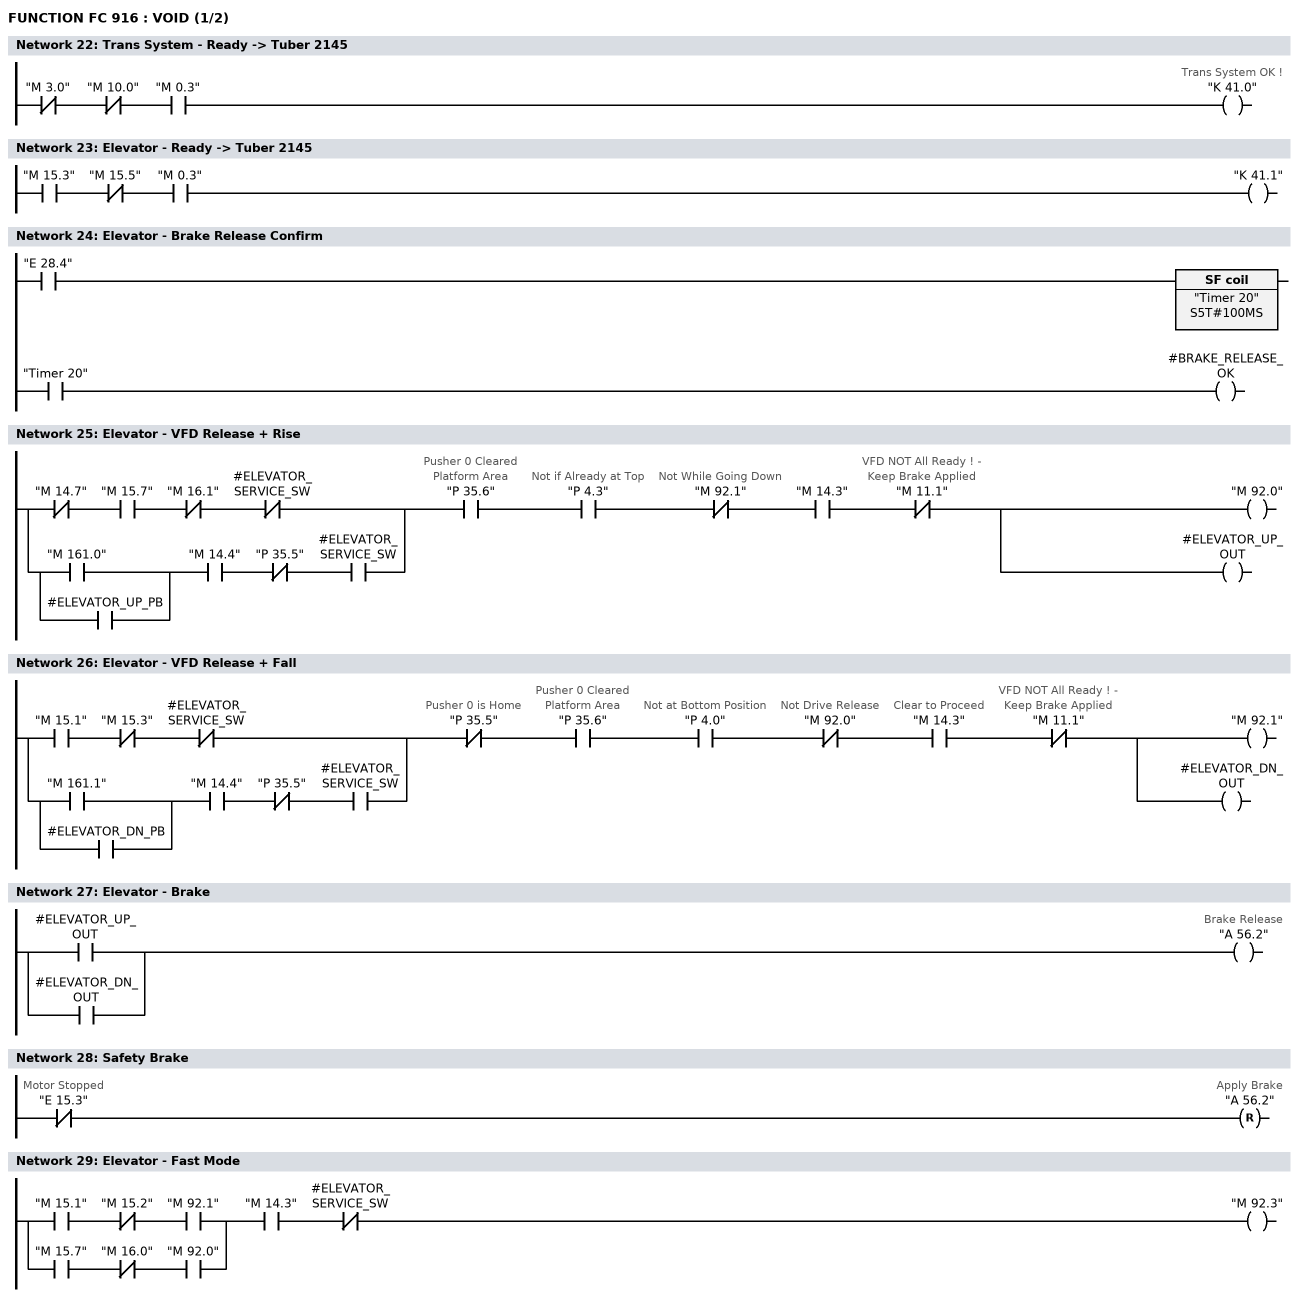

      AN    "M 3.0";
      AN    "M 10.0";
      A     "M 0.3";
      =     "K 41.0"; // Trans System OK !
NETWORK
TITLE =Elevator - Ready -> Tuber 2145

      A     "M 15.3";
      AN    "M 15.5";
      A     "M 0.3";
      =     "K 41.1";
NETWORK
TITLE =Elevator - Brake Release Confirm

      A     "E 28.4";
      L     S5T#100MS;
      SF    "Timer 20";
//;
      A     "Timer 20";
      =     #BRAKE_RELEASE_OK;
NETWORK
TITLE =Elevator - VFD Release + Rise

      A(    ;
      AN    "M 14.7";
      A     "M 15.7";
      AN    "M 16.1";
      AN    #ELEVATOR_SERVICE_SW;
      O     ;
      A(    ;
      O     "M 161.0";
      O     #ELEVATOR_UP_PB;
      )     ;
      A     "M 14.4";
      AN    "P 35.5";
      A     #ELEVATOR_SERVICE_SW;
      )     ;
      A     "P 35.6"; // Pusher 0 Cleared Platform Area
      A     "P 4.3"; // Not if Already at Top
      AN    "M 92.1"; // Not While Going Down
      A     "M 14.3";
      AN    "M 11.1"; // VFD NOT All Ready ! - Keep Brake Applied
      =     "M 92.0";
      =     #ELEVATOR_UP_OUT;
NETWORK
TITLE =Elevator - VFD Release + Fall

      A(    ;
      A     "M 15.1";
      AN    "M 15.3";
      AN    #ELEVATOR_SERVICE_SW;
      O     ;
      A(    ;
      O     "M 161.1";
      O     #ELEVATOR_DN_PB;
      )     ;
      A     "M 14.4";
      AN    "P 35.5";
      A     #ELEVATOR_SERVICE_SW;
      )     ;
      AN    "P 35.5"; // Pusher 0 is Home
      A     "P 35.6"; // Pusher 0 Cleared Platform Area
      A     "P 4.0"; // Not at Bottom Position
      AN    "M 92.0"; // Not Drive Release
      A     "M 14.3"; // Clear to Proceed
      AN    "M 11.1"; // VFD NOT All Ready ! - Keep Brake Applied
      =     "M 92.1";
      =     #ELEVATOR_DN_OUT;
NETWORK
TITLE =Elevator - Brake

      A(    ;
      O     #ELEVATOR_UP_OUT;
      O     #ELEVATOR_DN_OUT;
      )     ;
      =     "A 56.2"; // Brake Release
NETWORK
TITLE =Safety Brake

      AN    "E 15.3"; // Motor Stopped
      R     "A 56.2"; // Apply Brake
NETWORK
TITLE =Elevator - Fast Mode

      A(    ;
      A     "M 15.1";
      AN    "M 15.2";
      A     "M 92.1";
      O     ;
      A     "M 15.7";
      AN    "M 16.0";
      A     "M 92.0";
      )     ;
      A     "M 14.3";
      AN    #ELEVATOR_SERVICE_SW;
      =     "M 92.3";
NETWORK
TITLE =Elevator - Slow
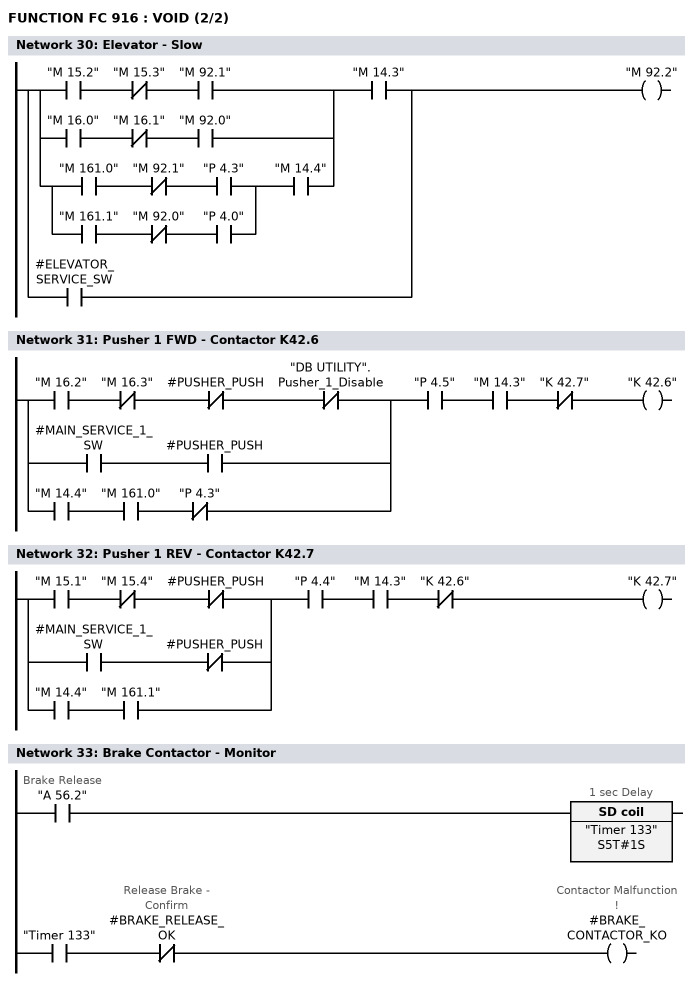

      A(    ;
      A     "M 15.2";
      AN    "M 15.3";
      A     "M 92.1";
      O     ;
      A     "M 16.0";
      AN    "M 16.1";
      A     "M 92.0";
      O     ;
      A(    ;
      A     "M 161.0";
      AN    "M 92.1";
      A     "P 4.3";
      O     ;
      A     "M 161.1";
      AN    "M 92.0";
      A     "P 4.0";
      )     ;
      A     "M 14.4";
      )     ;
      A     "M 14.3";
      O     #ELEVATOR_SERVICE_SW;
      =     "M 92.2";
NETWORK
TITLE =Pusher 1 FWD - Contactor K42.6

      A(    ;
      A     "M 16.2";
      AN    "M 16.3";
      AN    #PUSHER_PUSH;
      AN    "DB UTILITY".Pusher_1_Disable;
      O(    ;
      A     #MAIN_SERVICE_1_SW;
      A     #PUSHER_PUSH;
      )     ;
      O     ;
      A     "M 14.4";
      A     "M 161.0";
      AN    "P 4.3";
      )     ;
      A     "P 4.5";
      A     "M 14.3";
      AN    "K 42.7";
      =     "K 42.6";
NETWORK
TITLE =Pusher 1 REV - Contactor K42.7

      A(    ;
      A     "M 15.1";
      AN    "M 15.4";
      AN    #PUSHER_PUSH;
      O(    ;
      A     #MAIN_SERVICE_1_SW;
      AN    #PUSHER_PUSH;
      )     ;
      O     ;
      A     "M 14.4";
      A     "M 161.1";
      )     ;
      A     "P 4.4";
      A     "M 14.3";
      AN    "K 42.6";
      =     "K 42.7";
NETWORK
TITLE =Brake Contactor - Monitor

      A     "A 56.2"; // Brake Release
      L     S5T#1S; // 1 sec Delay
      SD    "Timer 133";
//;
      A     "Timer 133";
      AN    #BRAKE_RELEASE_OK; // Release Brake - Confirm
      =     #BRAKE_CONTACTOR_KO; // Contactor Malfunction !
NETWORK
TITLE =New Elevator VFD PARKER - Ready

      AN    "E 14.4"; // DRIVE TEST
      O     #BRAKE_CONTACTOR_KO; // Contactor Monitor = Contactor Malfunction !
      JCN   NFLT; // No fault
      S     "M 92.5"; // Set Fault Bit
      JU    OFF; // Turn Off
NETWORK
TITLE =New Elevator VFD with Dynamic Resistor - Go Up

NFLT: A     #ELEVATOR_UP_OUT; // VFD Release Command UP
      A     "M 92.3"; // Fast Speed Command
      AN    "M 92.5"; // Fault Bit
      AN    "M 11.1"; // VFD NOT All Ready !
      JCN   UPLO;
      S     "A 63.0"; // Release Drive - Go Up
      S     "A 63.2"; // Speed 2 / Speed 0.0
//;
      A     #BRAKE_RELEASE_OK; // Release Brake - Confirm
      JCN   END;
      =     "A 63.1"; // Speed 1
      =     "A 63.2"; // Speed 2 + Speed 1 = Fast
      R     "A 63.3"; // L = Forward (Up)
      JU    END;

UPLO: A     #ELEVATOR_UP_OUT; // VFD Release Command UP
      A     "M 92.2"; // Slow Speed Command
      AN    "M 92.5"; // Fault Bit
      AN    "M 11.1"; // VFD NOT All Ready !
      JCN   DNHI;
      S     "A 63.0"; // Release Drive - Go Up
      S     "A 63.2"; // Speed 2 / Speed 0.0
//;
      A     #BRAKE_RELEASE_OK; // Release Brake - Confirm
      JCN   END;
      =     "A 63.1"; // Speed 1
      R     "A 63.2"; // Speed 2 = Off
      R     "A 63.3"; // L = Forward (Up)
      JU    END;
NETWORK
TITLE =New Elevator VFD with Dynamic Resistor - Go Down

DNHI: A     #ELEVATOR_DN_OUT; // VFD Release Command DN
      A     "M 92.3"; // Fast Speed Command
      AN    "M 92.5"; // Fault Bit
      JCN   DNLO;
      S     "A 63.0"; // Release Drive - Go Dn
      S     "A 63.2"; // Speed 2 / Speed 0.0
//;
      A     #BRAKE_RELEASE_OK; // Release Brake - Confirm
      JCN   END;
      =     "A 63.1"; // Speed 1
      =     "A 63.2"; // Speed 2 + Speed 1 = Fast
      =     "A 63.3"; // H = Reverse (Dn)
      JU    END;

DNLO: A     #ELEVATOR_DN_OUT; // VFD Release Command DN
      A     "M 92.2"; // Slow Speed Command
      AN    "M 92.5"; // Fault Bit
      JCN   OFF;
      S     "A 63.0"; // Release Drive - Go Dn
      S     "A 63.2"; // Speed 2 / Speed 0.0
//;
      A     #BRAKE_RELEASE_OK; // Release Brake - Confirm
      JCN   END;
      =     "A 63.1"; // Speed 1
      R     "A 63.2"; // Speed 2 = Off
      =     "A 63.3"; // H = Reverse (Dn)
      JU    END;
NETWORK
TITLE =Drive Off
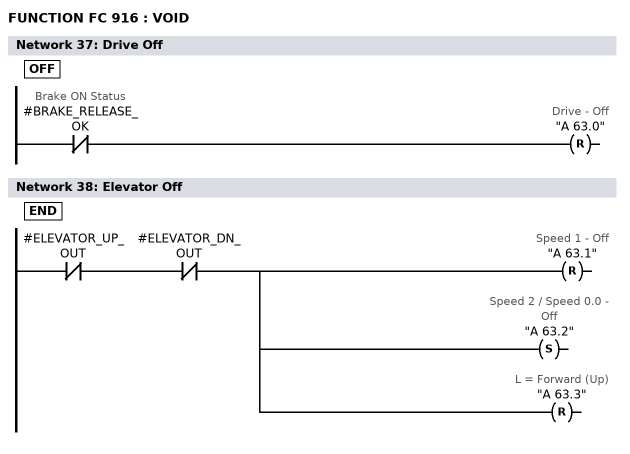

OFF:  AN    #BRAKE_RELEASE_OK; // Brake ON Status
      R     "A 63.0"; // Drive - Off
NETWORK
TITLE =Elevator Off

END:  AN    #ELEVATOR_UP_OUT;
      AN    #ELEVATOR_DN_OUT;
      R     "A 63.1"; // Speed 1 - Off
      S     "A 63.2"; // Speed 2 / Speed 0.0 - Off
      R     "A 63.3"; // L = Forward (Up)
END_FUNCTION


FUNCTION FC 918 : VOID
TITLE =NEW FC918 (was FC1018) - Conveyor 1 Pos. 1
//
NAME : POS_3
VERSION : 0.0


VAR_TEMP
  MAIN_SERVICE_1_SW : BOOL ;
  SERVICE_RUN : BOOL ;
  INITIALISATION : BOOL ;
  SENSOR_TEST : BOOL ;
END_VAR
BEGIN
NETWORK
TITLE =Service Test

      A     "HMI_DB".ALL_SERVICE_ENABLE_SW;
      A     "HMI_DB".CONVEYOR_1_SERVICE_SW;
      A     "HMI_DB".SERVICE_SW_1_STATUS;
      =     #MAIN_SERVICE_1_SW;
//;
      A     #MAIN_SERVICE_1_SW;
      O     "M 18.1";
      JNB   CON1;
      A     "HMI_DB".HMI_CONVEYOR_1_TEST_SSW;
      =     #SERVICE_RUN;
      S     "DB UTILITY".Elevator_Disable;
      S     "DB UTILITY".Pusher_1_Disable;
//;
      A     "HMI_DB".SERVICE_INIT_PB;
      =     #INITIALISATION;
//;
      AN    #MAIN_SERVICE_1_SW;
      R     "HMI_DB".HMI_CONVEYOR_1_TEST_SSW;
      R     "DB UTILITY".Elevator_Disable;
      R     "DB UTILITY".Pusher_1_Disable;

CON1: R     #SERVICE_RUN;
      R     #INITIALISATION;
      FP    "FP 158.2";
      =     "M 18.1";
NETWORK
TITLE =Step 2N1 - Power ON
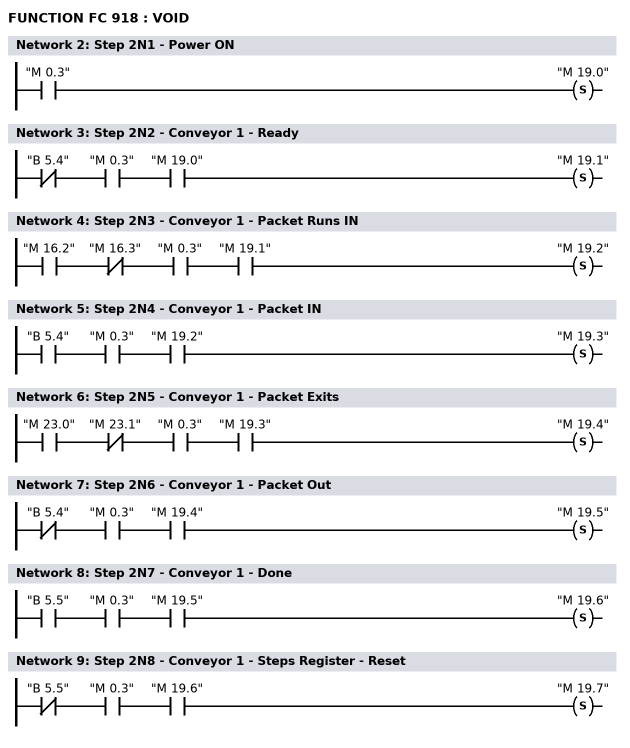

      A     "M 0.3";
      S     "M 19.0";
NETWORK
TITLE =Step 2N2 - Conveyor 1 - Ready

      AN    "B 5.4";
      A     "M 0.3";
      A     "M 19.0";
      S     "M 19.1";
NETWORK
TITLE =Step 2N3 - Conveyor 1 - Packet Runs IN

      A     "M 16.2";
      AN    "M 16.3";
      A     "M 0.3";
      A     "M 19.1";
      S     "M 19.2";
NETWORK
TITLE =Step 2N4 - Conveyor 1 - Packet IN

      A     "B 5.4";
      A     "M 0.3";
      A     "M 19.2";
      S     "M 19.3";
NETWORK
TITLE =Step 2N5 - Conveyor 1 - Packet Exits

      A     "M 23.0";
      AN    "M 23.1";
      A     "M 0.3";
      A     "M 19.3";
      S     "M 19.4";
NETWORK
TITLE =Step 2N6 - Conveyor 1 - Packet Out

      AN    "B 5.4";
      A     "M 0.3";
      A     "M 19.4";
      S     "M 19.5";
NETWORK
TITLE =Step 2N7 - Conveyor 1 - Done

      A     "B 5.5";
      A     "M 0.3";
      A     "M 19.5";
      S     "M 19.6";
NETWORK
TITLE =Step 2N8 - Conveyor 1 - Steps Register - Reset

      AN    "B 5.5";
      A     "M 0.3";
      A     "M 19.6";
      S     "M 19.7";
NETWORK
TITLE =Conveyor 1 - Steps Register - Reset

      A(    ;
      O     "M 19.7";
      O     "DB UTILITY".T19_DN;
      O     #INITIALISATION;
      O     "DB UTILITY".Conveyor_1_Disable;
      )     ;
      A     "M 0.3";
      JNB   INIT;
      L     W#16#0;
      T     "MW 19";

INIT: CLR   ;
NETWORK
TITLE =Soft Timer 19 Reset

      A     "M 19.2";
      AN    "M 19.3";
      A     "M 0.3";
      JCN   R191;
      JU    E191;

R191: L     L#0;
      T     "DB UTILITY".T19_ET;
      R     "DB UTILITY".T19_DN;

E191: NOP   0;

NETWORK
TITLE =Soft Timer 19 Add

      A     "M 19.2";
      AN    "M 19.3";
      A     "M 0.3";
      AN    "DB UTILITY".Freeze_Sequence_1;
      AN    "DB UTILITY".T19_DN;
      JCN   E192;

      L     "DB UTILITY".T19_ET;
      L     "DB UTILITY".Scan_Cycle_Previous;
      ITD   ;
      +D    ;
      T     "DB UTILITY".T19_ET;

E192: NOP   0;

NETWORK
TITLE =Soft Timer 19 Done 10s
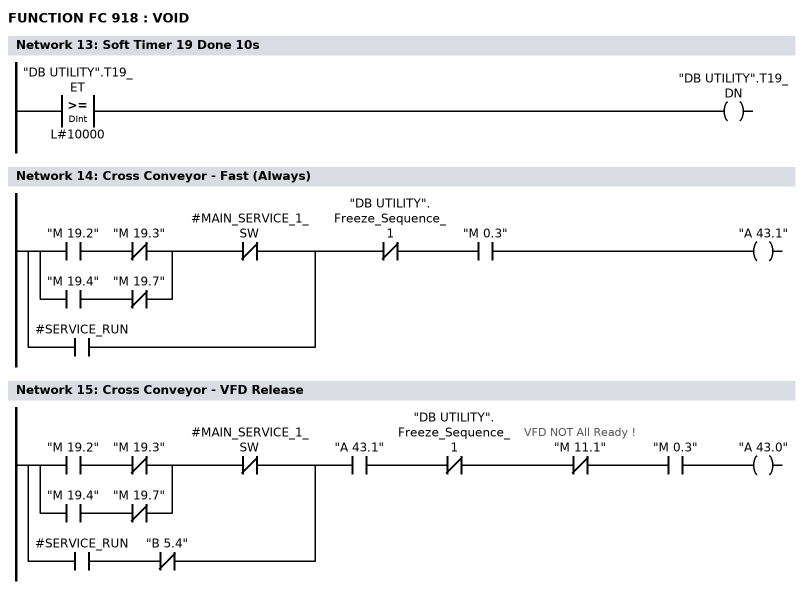

      L     "DB UTILITY".T19_ET;
      L     L#10000;
      >=D   ;
      =     "DB UTILITY".T19_DN;
NETWORK
TITLE =Cross Conveyor - Fast (Always)

      A(    ;
      A     "M 19.2";
      AN    "M 19.3";
      O     ;
      A     "M 19.4";
      AN    "M 19.7";
      )     ;
      AN    #MAIN_SERVICE_1_SW;
      O     #SERVICE_RUN;
      AN    "DB UTILITY".Freeze_Sequence_1;
      A     "M 0.3";
      =     "A 43.1";

NETWORK
TITLE =Cross Conveyor - VFD Release

      A(    ;
      A     "M 19.2";
      AN    "M 19.3";
      O     ;
      A     "M 19.4";
      AN    "M 19.7";
      )     ;
      AN    #MAIN_SERVICE_1_SW;
      O(    ;
      A     #SERVICE_RUN;
      AN    "B 5.4";
      )     ;
      A     "A 43.1";
      AN    "DB UTILITY".Freeze_Sequence_1;
      AN    "M 11.1"; // VFD NOT All Ready !
      A     "M 0.3";
      =     "A 43.0";
NETWORK
TITLE =Any Conveyors Packet mS Test

//    A     "B 10.7"
//    A     "A 48.6"


      A     "B 10.6";
      A     "A 48.3";






      =     #SENSOR_TEST;
//;
      A     #SENSOR_TEST;
      FP    "FP 147.7";
      JNB   NRST;
      L     0;
      T     "COLLATORS DB".Any_Conveyors_mS;

NRST: A     #SENSOR_TEST;
      JNB   NCNT;
      L     "COLLATORS DB".Any_Conveyors_mS;
      L     "DB UTILITY".Scan_Cycle_Previous;
      ITD   ;
      +D    ;
      T     "COLLATORS DB".Any_Conveyors_mS;

NCNT: CLR   ;

END_FUNCTION


FUNCTION FC 922 : VOID
TITLE =NEW FC922 (was FC1022) - Angle Conveyor 2 Pos. 4
NAME : POS_4
VERSION : 0.0


VAR_TEMP
  MAIN_SERVICE_1_SW : BOOL ;
  SERVICE_BELT_RUN : BOOL ;
  SERVICE_ROLLER_LIFT : BOOL ;
  SERVICE_ROLLER_RUN : BOOL ;
  INITIALISATION : BOOL ;
  PACKET_MEASURE_FLAG : BOOL ;
END_VAR
BEGIN
NETWORK
TITLE =Service Test

      A     "HMI_DB".ALL_SERVICE_ENABLE_SW;
      A     "HMI_DB".CONVEYOR_2_SERVICE_SW;
      A     "HMI_DB".SERVICE_SW_1_STATUS;
      =     #MAIN_SERVICE_1_SW;
//;
      A     #MAIN_SERVICE_1_SW;
      O     "M 22.1";
      JNB   CON2;
      A     "HMI_DB".HMI_CONVEYOR_2B_TEST_SSW;
      =     #SERVICE_BELT_RUN;
      S     "DB UTILITY".Conveyor_1_Disable;
//;
      A     "HMI_DB".HMI_CONVEYOR_2L_TEST_SSW;
      =     #SERVICE_ROLLER_LIFT;
      S     "DB UTILITY".Conveyor_1_Disable;
//;
      A     "HMI_DB".HMI_CONVEYOR_2R_TEST_SSW;
      =     #SERVICE_ROLLER_RUN;
      S     "DB UTILITY".Conveyor_1_Disable;
//;
      A     "HMI_DB".SERVICE_INIT_PB;
      =     #INITIALISATION;
//;
      AN    #MAIN_SERVICE_1_SW;
      R     "HMI_DB".HMI_CONVEYOR_2B_TEST_SSW;
      R     "HMI_DB".HMI_CONVEYOR_2L_TEST_SSW;
      R     "HMI_DB".HMI_CONVEYOR_2R_TEST_SSW;
      R     "DB UTILITY".Conveyor_1_Disable;

CON2: R     #SERVICE_BELT_RUN;
      R     #SERVICE_ROLLER_LIFT;
      R     #SERVICE_ROLLER_RUN;
      R     #INITIALISATION;
      FP    "FP 158.3";
      =     "M 22.1";

NETWORK
TITLE =Angle Conveyor - Fault / Ready
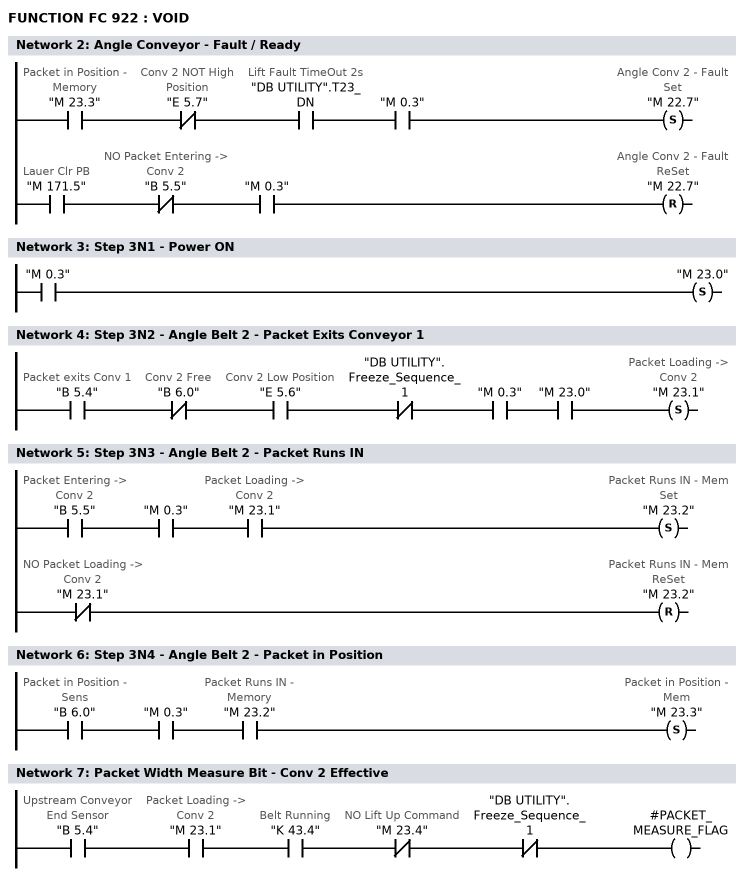

      A     "M 23.3"; // Packet in Position - Memory
      AN    "E 5.7"; // Conv 2 NOT High Position
      A     "DB UTILITY".T23_DN; // Lift Fault TimeOut 2s
      A     "M 0.3";
      S     "M 22.7"; // Angle Conv 2 - Fault Set
//;
      A     "M 171.5"; // Lauer Clr PB
      AN    "B 5.5"; // NO Packet Entering -> Conv 2
      A     "M 0.3";
      R     "M 22.7"; // Angle Conv 2 - Fault ReSet

NETWORK
TITLE =Step 3N1 - Power ON

      A     "M 0.3";
      S     "M 23.0";

NETWORK
TITLE =Step 3N2 - Angle Belt 2 - Packet Exits Conveyor 1

      A     "B 5.4"; // Packet exits Conv 1
      AN    "B 6.0"; // Conv 2 Free
      A     "E 5.6"; // Conv 2 Low Position
      AN    "DB UTILITY".Freeze_Sequence_1;
      A     "M 0.3";
      A     "M 23.0";
      S     "M 23.1"; // Packet Loading -> Conv 2
NETWORK
TITLE =Step 3N3 - Angle Belt 2 - Packet Runs IN

      A     "B 5.5"; // Packet Entering -> Conv 2
      A     "M 0.3";
      A     "M 23.1"; // Packet Loading -> Conv 2
      S     "M 23.2"; // Packet Runs IN - Mem Set
//;
      ON    "M 23.1"; // NO Packet Loading -> Conv 2
      R     "M 23.2"; // Packet Runs IN - Mem ReSet

NETWORK
TITLE =Step 3N4 - Angle Belt 2 - Packet in Position

      A     "B 6.0"; // Packet in Position - Sens
      A     "M 0.3";
      A     "M 23.2"; // Packet Runs IN - Memory
      S     "M 23.3"; // Packet in Position - Mem
NETWORK
TITLE =Packet Width Measure Bit - Conv 2 Effective

      A     "B 5.4"; // Upstream Conveyor End Sensor
      A     "M 23.1"; // Packet Loading -> Conv 2
      A     "K 43.4"; // Belt Running
      AN    "M 23.4"; // NO Lift Up Command
      AN    "DB UTILITY".Freeze_Sequence_1;
      =     #PACKET_MEASURE_FLAG;

NETWORK
TITLE =Packet Width Time Reset - Freeze Safe

      A     "M 23.1"; // Packet Loading -> Conv 2
      O     "DB UTILITY".Freeze_Sequence_1;
      JC    NRS1;

      L     L#0;
      T     "MD 260"; // Width [mS]

NRS1: NOP   0;
NETWORK
TITLE =Packet Width Time Count Up From Sensor "B 5.4"

      A     #PACKET_MEASURE_FLAG;
      JCN   NMES;

      L     "MD 260"; // Width [mS]
      L     "DB UTILITY".Scan_Cycle_Previous;
      ITD   ;
      +D    ;
      T     "MD 260"; // Width [mS]

NMES: NOP   0;
NETWORK
TITLE =Middle Travel Time Reset - Freeze Safe

      A     "M 23.3"; // Packet in Position - Mem
      O     "DB UTILITY".Freeze_Sequence_1;
      JC    NRS2;

      L     L#0;
      T     "MD 264"; // Half Width [mS] - Zeroed

NRS2: NOP   0;
NETWORK
TITLE =Middle Travel Time Count Up From B 6.0

      ON    "M 23.3"; // NO Packet in Position - Mem
      O     "M 23.4"; // Lift Up Command
      ON    "K 43.4"; // Belt Stopped
      ON    "M 0.3"; // No Power
      AN    "DB UTILITY".Freeze_Sequence_1;
      JC    NCNT;

      L     "MD 264"; // Half Width [mS]
      L     "DB UTILITY".Scan_Cycle_Previous;
      ITD   ;
      +D    ;
      T     "MD 264"; // Half Width [mS] - Add

NCNT: NOP   0;
NETWORK
TITLE =Middle Travel Time Clamp Zero

      L     "MD 264"; // Half Width [mS]
      L     L#0;
      >=D   ;
      JC    NMID;

      L     L#0;
      T     "MD 264"; // Half Width [mS] - Reset

NMID: NOP   0;
NETWORK
TITLE =Soft Timer 23 Reset - Lift Fault TimeOut 2s + Freeze Option

      A     "M 23.3"; // Packet in Position - Memory
      AN    "M 23.4"; // NO Lift Up Command
      A     "M 0.3";
      JCN   R231;
      JU    E231;

R231: L     L#0;
      T     "DB UTILITY".T23_ET;
      R     "DB UTILITY".T23_DN;

E231: NOP   0;

NETWORK
TITLE =Soft Timer 23 Add

      A     "M 23.3"; // Packet in Position - Memory
      AN    "M 23.4"; // NO Lift Up Command
      A     "M 0.3";
      AN    "DB UTILITY".Freeze_Sequence_1; // Sequence Freezer Bit
      AN    "DB UTILITY".T23_DN;
      JCN   E232;

      L     "DB UTILITY".T23_ET;
      L     "DB UTILITY".Scan_Cycle_Previous;
      ITD   ;
      +D    ;
      T     "DB UTILITY".T23_ET;

E232: NOP   0;

NETWORK
TITLE =Soft Timer 23 Done 2s

      L     "DB UTILITY".T23_ET;
      L     L#2500; // [mS]
      >=D   ;
      =     "DB UTILITY".T23_DN;
NETWORK
TITLE =Soft Timer 24 Reset - Belt TimeOut 8s + Freeze Option

      A     "M 23.1";
      AN    "M 23.3";
      A     "K 43.4";
      A     "M 0.3";
      JCN   R241;
      JU    E241;

R241: L     L#0;
      T     "DB UTILITY".T24_ET;
      R     "DB UTILITY".T24_DN;

E241: NOP   0;

NETWORK
TITLE =Soft Timer 24 Add

      A     "M 23.1";
      AN    "M 23.3";
      A     "K 43.4";
      A     "M 0.3";
      AN    "DB UTILITY".Freeze_Sequence_1;
      AN    "DB UTILITY".T24_DN;
      JCN   E242;

      L     "DB UTILITY".T24_ET;
      L     "DB UTILITY".Scan_Cycle_Previous;
      ITD   ;
      +D    ;
      T     "DB UTILITY".T24_ET;

E242: NOP   0;

NETWORK
TITLE =Soft Timer 24 Done 8s

      L     "DB UTILITY".T24_ET;
      L     L#8000;
      >=D   ;
      =     "DB UTILITY".T24_DN;
      S     "M 24.4";
NETWORK
TITLE =Step 3N5 - Angle Belt - Lift ("MD 264" to Center the Packet)

      A(    ;
      A(    ;
      L     "MD 264";
      L     L#2;
      *D    ;
      L     "MD 260";
      >=D   ;
      )     ;
      AN    #PACKET_MEASURE_FLAG;
      AN    "B 5.5";
      O     "DB UTILITY".T23_DN;
      )     ;
      A     "M 0.3";
      A     "M 23.3";
      S     "M 23.4";
NETWORK
TITLE =Step 3N6 - Angle Rollers - Up
